(* IEC 61131-3 sources: daoli-st-library/DL_Process (part 36) *)

(* ---- FB_DL_GrateCoolerStartupSeq.st ---- *)
(*
  Name: FB_DL_GrateCoolerStartupSeq
  Category: DL_Process
  Version: 1.0.0
  Round: R91 / 2026-11-25
  开源溯源：clean-room 自研（族 水泥窑篦冷机与预热器，ST 开源生态实测 0 命中，无外部代码引入）
  功能：1) 篦冷机启动序状态机，七相推进：
           待机 → 风机启动 → 篦床低速 → 投料 → 投料升速 → 正常 → （故障）。
           待机相等 xStart 上升沿（必须边沿，防上电即在启动位自动启动）；
           风机相开风机命令并等运行反馈 + 风量达启动下限；篦床低速相给低速指令并等运行反馈；
           投料相开投料命令并等投料反馈；升速相把转速指令按 fRampRpmS 斜率从低速升到正常；
           正常相保持 xDone 并继续风量安全监督，直到 xStart 撤下才回待机。
        2) 每相独立超时 + 整序总超时：相定时器给出正常推进点，相超时定时器给出
           「定时 + DL_OVER_MARGIN」的越限点，整序总超时由 tonTotal 兜底，三者并发监视。
        3) 风量安全监督分两段语义：启动阶段风量不足只拦放行并置信息级码（0121），
           投料之后风量跌破安全下限则进入宽限窗，宽限超时判故障（0128，防篦板过热）。
  边界条件：1) 非有限值闸：风量、转速反馈、周期入参先过 NOT(x > -DL_BIG AND x < DL_BIG)，
           同时拦 NaN 与 Inf；命中即闸断放行（_bAirOk := FALSE / 停机相），
           绝不把 NaN 与 DL_AIR_MIN 比较 —— NaN 比较恒假会伪装成「风量正常」（R19）。
        2) 周期入参闸（R21）：fCycleS <= 0.0 或非有限时，一律改用缺省 DL_CYCLE_DEF = 0.1 s，
           并置信息级码 0129 声明本次斜率按缺省周期折算，不静默。
        3) 时间参数零闸：tFanS / tGrateS / tFeedS / tRampS <= T#0S 时对应相定时器立即置 Q，
           等价于该相跳过（调试用合法组态），语义在此声明，禁上层按「必有停留」假设。
        4) 斜率上限：升速相每拍增量 = fRampRpmS * fCycleS，且指令本身钳在
           [DL_SPD_SLOW, DL_SPD_NORMAL] 内，不用 LIMIT 之后再判超限（R24）。
        5) 故障归因唯一（R190）：风机超时 / 篦床超时 / 投料超时 / 升速超时 / 总超时 /
           外部故障 / 风量不足 / 兜底，八条成因各占独立码值，不共用枚举成员。
        6) 故障解除路径：故障相内 xReset 上升沿 AND NOT xFault AND 入参有限 → 清锁存回待机；
           回待机后必须重新给 xStart 上升沿才能再启动（不自恢复）。
        7) 状态机兜底：CASE 全态覆盖 + ELSE 强制回故障相并置码 0130、清全部输出。
        8) 输出安全初值（R25）：fGrateSpdCmdRpm 初值 0.0（零速为安全侧），
           三个命令位初值 FALSE，待机相显式赋值，防「上电 0 值直穿下发」。
  量纲自证：fRampRpmS 为转速斜率 [rpm/s]，乘 fCycleS [s] 得每拍增量 [rpm]，
           与 fGrateSpdCmdRpm [rpm] 同量纲；fAirFlowNm3h 与 DL_AIR_MIN 同量纲 [Nm3/h]；
           所有时间引脚为 [TIME]，相超时点 = [TIME] + [TIME] = [TIME]，与 TON 的 PT 同量纲。
  码表 Error codes（本件子带 0091_012x，故障级一律 3 行内置 _uFault/_bFault/_eState）:
    16#0091_0121 信息级：风量低于启动下限，风机相暂不放行（不置故障位）
    16#0091_0122 故障级：风机启动超时（定时到但运行反馈未到）
    16#0091_0123 故障级：篦床低速启动超时（无运行反馈）
    16#0091_0124 故障级：投料超时（无投料反馈）
    16#0091_0125 故障级：升速超时（未达正常转速）
    16#0091_0126 故障级：整序总超时
    16#0091_0127 故障级：外部故障输入 xFault
    16#0091_0128 故障级：运行中风量低于安全下限（宽限窗超时）
    16#0091_0129 信息级：周期入参 fCycleS 非法，已按缺省 0.1 s 折算（不置故障位）
    16#0091_0130 故障级：状态机落 ELSE 兜底（非法相位 ID）
    16#0091_0131 故障级：启动序期间风量/转速/斜率入参非有限（NaN 或 Inf）

  修订历史 Revision :
    2026-11-25  v1.0.0  R91 首版
*)

TYPE E_DL_GcsStartupState :
(
    eGcsStartIdle      := 0,    // 待机：等启动上升沿 / Idle, awaiting the start rising edge
    eGcsStartFan       := 10,   // 风机启动：等运行反馈与风量 / Fan start, awaiting feedback and air flow
    eGcsStartSlowGrate := 20,   // 篦床低速：给低速指令等运行反馈 / Grate at low speed, awaiting run feedback
    eGcsStartFeed      := 30,   // 投料：开投料命令等投料反馈 / Feeding, awaiting the feed feedback
    eGcsStartRampUp    := 40,   // 投料升速：按斜率升到正常转速 / Ramping up to normal speed
    eGcsStartNormal    := 50,   // 正常：保持完成位并继续风量监督 / Normal, done held and air supervised
    eGcsStartFault     := 90    // 故障：锁存待解除 / Fault, latched awaiting release
);
END_TYPE

FUNCTION_BLOCK FB_DL_GrateCoolerStartupSeq
VAR_INPUT
    xStart        : BOOL;    // 启动指令（上升沿有效）[bool] / Start command, edge triggered [bool]
    xReset        : BOOL;    // 故障复位（上升沿有效）[bool] / Fault reset, rising edge [bool]
    xFault        : BOOL;    // 外部故障汇总 [bool] / External fault aggregate [bool]
    xFanRunFb     : BOOL;    // 风机运行反馈 [bool] / Fan running feedback [bool]
    xGrateRunFb   : BOOL;    // 篦床驱动运行反馈 [bool] / Grate drive running feedback [bool]
    xFeedRunFb    : BOOL;    // 投料设备运行反馈 [bool] / Feed device running feedback [bool]
    fAirFlowNm3h  : REAL;    // 冷却风量实测值 [Nm3/h] / Measured cooling air flow [Nm3/h]
    fGrateSpdFbRpm : REAL;   // 篦床转速反馈 [rpm] / Grate speed feedback [rpm]
    fRampRpmS     : REAL;    // 升速斜率 [rpm/s] / Speed ramp slope [rpm/s]
    fCycleS       : REAL;    // 任务周期 [s] / Task cycle time [s]
    tFanS         : TIME;    // 风机相设定时长 [TIME] / Fan phase duration [TIME]
    tGrateS       : TIME;    // 篦床低速相设定时长 [TIME] / Low-speed grate phase duration [TIME]
    tFeedS        : TIME;    // 投料相设定时长 [TIME] / Feeding phase duration [TIME]
    tRampS        : TIME;    // 升速相设定时长 [TIME] / Ramp-up phase duration [TIME]
END_VAR
VAR_OUTPUT
    xFanCmd       : BOOL;    // 风机运行命令（安全侧：故障时停）[bool] / Fan run command, fail-safe [bool]
    xGrateCmd     : BOOL;    // 篦床驱动运行命令（安全侧：故障时停）[bool] / Grate drive command, fail-safe [bool]
    xFeedCmd      : BOOL;    // 投料设备运行命令（安全侧：故障时停）[bool] / Feed device command, fail-safe [bool]
    fGrateSpdCmdRpm : REAL;  // 篦床转速指令 [rpm] / Grate speed command [rpm]
    xDone         : BOOL;    // 启动完成保持位 [bool] / Startup complete held flag [bool]
    xBusy         : BOOL;    // 启动进行中 [bool] / Startup sequence busy [bool]
    xAirOk        : BOOL;    // 风量监督通过 [bool] / Air flow supervision passed [bool]
    eState        : E_DL_GcsStartupState;   // 状态出口，段尾单点映射 / State outlet, single-point mapped
    nErrId        : UDINT;   // 事件码，0 = 无事件 / Event code, 0 = none
END_VAR
VAR
    tonFan        : TON;     // 风机相正常定时 [TIME] / Fan phase timer
    tonFanOv      : TON;     // 风机相超时定时 [TIME] / Fan phase overrun timer
    tonGrate      : TON;     // 篦床低速相正常定时 [TIME] / Low-speed grate phase timer
    tonGrateOv    : TON;     // 篦床低速相超时定时 [TIME] / Low-speed grate phase overrun timer
    tonFeed       : TON;     // 投料相正常定时 [TIME] / Feeding phase timer
    tonFeedOv     : TON;     // 投料相超时定时 [TIME] / Feeding phase overrun timer
    tonRamp       : TON;     // 升速相正常定时 [TIME] / Ramp-up phase timer
    tonRampOv     : TON;     // 升速相超时定时 [TIME] / Ramp-up phase overrun timer
    tonTotal      : TON;     // 整序总超时定时 [TIME] / Whole-sequence total timeout timer
    tonAirG       : TON;     // 运行中风量不足宽限定时 [TIME] / Air-shortage grace timer while running
    rtStart       : R_TRIG;  // 启动上升沿检测 [bool] / Start rising edge detector
    rtReset       : R_TRIG;  // 复位上升沿检测 [bool] / Reset rising edge detector
    _eState       : E_DL_GcsStartupState := E_DL_GcsStartupState.eGcsStartIdle;   // 内部相位（CASE 唯一写入目标）
    _eStatePrev   : E_DL_GcsStartupState := E_DL_GcsStartupState.eGcsStartIdle;   // 上一拍相位快照（周期末更新）
    _fSpdSet      : REAL := 0.0;    // 转速指令内部设定值（安全初值零速）[rpm] / Internal speed setpoint, safe init zero [rpm]
    _fCycleUseS   : REAL := 0.1;    // 实际使用的周期值 [s] / Cycle time actually used [s]
    _bFinOk       : BOOL := FALSE;  // 实值入参有限性总闸结果 / Finiteness gate aggregate result
    _bCycleBad    : BOOL := FALSE;  // 周期入参非法标志 [bool] / Cycle input invalid flag [bool]
    _bAirOk       : BOOL := FALSE;  // 风量监督结果 [bool] / Air flow supervision result [bool]
    _bActive      : BOOL := FALSE;  // 启动序激活（风机至正常五相之一）[bool] / Sequence active flag [bool]
    _bRunAirWatch : BOOL := FALSE;  // 投料后风量安全监督生效 [bool] / Post-feed air supervision active [bool]
    _bDoneL       : BOOL := FALSE;  // 完成位锁存（跨相保持）[bool] / Done latch held across phases [bool]
    _bFault       : BOOL := FALSE;  // 故障锁存位 [bool] / Latched fault flag [bool]
    _bRampDone    : BOOL := FALSE;  // 升速到位标志（指令达正常转速）[bool] / Ramp-complete flag [bool]
    _uInfo        : UDINT := 16#0000_0000;   // 信息码，每拍重算 / Info code, recomputed every cycle
    _uFault       : UDINT := 16#0000_0000;   // 故障码锁存 / Latched fault code
    _iPhaseChg    : INT := 0;       // 本拍相位切换计数（观测用）[-] / Phase-change count this cycle [-]
END_VAR
VAR CONSTANT
    DL_EPS        : REAL := 1.0E-9;      // 数值零闸阈值 [-] / Numeric zero gate threshold [-]
    DL_BIG        : REAL := 1.0E12;      // 非有限值闸量级上限 [-] / Finiteness gate magnitude [-]
    DL_CYCLE_DEF  : REAL := 0.1;         // 缺省任务周期 [s] / Default task cycle time [s]
    DL_CYCLE_MIN  : REAL := 0.001;       // 周期合理下限 [s] / Cycle time reasonable low bound [s]
    DL_CYCLE_MAX  : REAL := 10.0;        // 周期合理上限 [s] / Cycle time reasonable high bound [s]
    DL_AIR_MIN    : REAL := 5000.0;      // 启动风量下限 [Nm3/h] / Air flow low limit for start [Nm3/h]
    DL_AIR_SAFE   : REAL := 3000.0;      // 运行风量安全下限 [Nm3/h] / Air flow safety low limit while running [Nm3/h]
    DL_SPD_SLOW   : REAL := 2.0;         // 篦床低速设定 [rpm] / Grate low speed setpoint [rpm]
    DL_SPD_NORMAL : REAL := 12.0;        // 篦床正常转速设定 [rpm] / Grate normal speed setpoint [rpm]
    DL_OVER_MARGIN : TIME := T#30S;      // 相超时相对正常定时的裕量 [TIME] / Phase overrun margin [TIME]
    DL_TOTAL_MAX  : TIME := T#30M;       // 整序总超时上限 [TIME] / Whole-sequence total timeout [TIME]
    DL_AIR_GRACE  : TIME := T#15S;       // 运行中风量不足宽限窗 [TIME] / Air-shortage grace window [TIME]
END_VAR

(* —— 段 0：单拍量预清零（锁存量 _uFault/_bFault/_bDoneL/_eStatePrev 不入清单，R187①） —— *)
_uInfo := 16#0000_0000;                     // 信息码每拍重算 / Info code recomputed
_iPhaseChg := 0;                            // 相位切换计数每拍重算 / Phase-change counter recomputed
nErrId := 16#0000_0000;                     // 事件码缺省无事件 / Event code defaults to none

(* —— 段 1：周期入参闸（R21：非法周期不静默，改用缺省并置信息码） —— *)
_bCycleBad := NOT (fCycleS > -DL_BIG AND fCycleS < DL_BIG)
              OR (fCycleS < DL_CYCLE_MIN) OR (fCycleS > DL_CYCLE_MAX);
IF _bCycleBad THEN
    _fCycleUseS := DL_CYCLE_DEF;            // 非法周期一律用缺省 0.1 s
    _uInfo := 16#0091_0129;                 // 信息级：周期入参非法，已用缺省（不置故障位）
ELSE
    _fCycleUseS := fCycleS;                 // 合法周期原值使用
END_IF

(* —— 段 2：非有限值闸（R19：闸断实值通路，风量/转速/斜率任一非有限即拒绝放行） —— *)
_bFinOk := (fAirFlowNm3h > -DL_BIG) AND (fAirFlowNm3h < DL_BIG)
           AND (fGrateSpdFbRpm > -DL_BIG) AND (fGrateSpdFbRpm < DL_BIG)
           AND (fRampRpmS > -DL_BIG) AND (fRampRpmS < DL_BIG);

(* —— 段 3：风量监督（启动用下限；非有限值直接判不通过，不参与比较） —— *)
IF NOT _bFinOk THEN
    _bAirOk := FALSE;                       // 非有限一律判不通过（安全侧）
ELSE
    _bAirOk := (fAirFlowNm3h >= DL_AIR_MIN);
END_IF

(* —— 段 4：状态派生量（本拍相位为上一拍末值，标准 FB 周期语义） —— *)
_bActive := (_eState = E_DL_GcsStartupState.eGcsStartFan)
            OR (_eState = E_DL_GcsStartupState.eGcsStartSlowGrate)
            OR (_eState = E_DL_GcsStartupState.eGcsStartFeed)
            OR (_eState = E_DL_GcsStartupState.eGcsStartRampUp)
            OR (_eState = E_DL_GcsStartupState.eGcsStartNormal);
_bRunAirWatch := (_eState = E_DL_GcsStartupState.eGcsStartFeed)
                 OR (_eState = E_DL_GcsStartupState.eGcsStartRampUp)
                 OR (_eState = E_DL_GcsStartupState.eGcsStartNormal);

(* —— 段 5：定时器与边沿无条件周期刷新（R7：调用语句不得置于 IF/CASE 内） —— *)
rtStart(CLK := xStart);                                                                 // 启动上升沿，每拍必调
rtReset(CLK := xReset);                                                                 // 复位上升沿，每拍必调
tonFan(IN := (_eState = E_DL_GcsStartupState.eGcsStartFan), PT := tFanS);               // 风机相正常定时
tonFanOv(IN := (_eState = E_DL_GcsStartupState.eGcsStartFan), PT := tFanS + DL_OVER_MARGIN);      // 风机相超时点
tonGrate(IN := (_eState = E_DL_GcsStartupState.eGcsStartSlowGrate), PT := tGrateS);     // 篦床低速相正常定时
tonGrateOv(IN := (_eState = E_DL_GcsStartupState.eGcsStartSlowGrate),
           PT := tGrateS + DL_OVER_MARGIN);                                             // 篦床低速相超时点
tonFeed(IN := (_eState = E_DL_GcsStartupState.eGcsStartFeed), PT := tFeedS);            // 投料相正常定时
tonFeedOv(IN := (_eState = E_DL_GcsStartupState.eGcsStartFeed), PT := tFeedS + DL_OVER_MARGIN);   // 投料相超时点
tonRamp(IN := (_eState = E_DL_GcsStartupState.eGcsStartRampUp), PT := tRampS);          // 升速相正常定时
tonRampOv(IN := (_eState = E_DL_GcsStartupState.eGcsStartRampUp), PT := tRampS + DL_OVER_MARGIN); // 升速相超时点
tonTotal(IN := _bActive, PT := DL_TOTAL_MAX);                                           // 整序总超时
tonAirG(IN := _bRunAirWatch AND (NOT _bAirOk) AND (NOT _bFault), PT := DL_AIR_GRACE);    // 风量不足宽限窗

(* —— 段 6：全局故障拦截（优先级最高；已锁存则不再改写码值，禁同拍抹除） —— *)
IF xFault AND (NOT _bFault) THEN
    _uFault := 16#0091_0127;                // 故障级：外部故障输入
    _bFault := TRUE;                        // 锁存（3 行内置，R45 配对）
    _eState := E_DL_GcsStartupState.eGcsStartFault;
END_IF
IF tonTotal.Q AND _bActive AND (NOT _bFault) THEN
    _uFault := 16#0091_0126;                // 故障级：整序总超时
    _bFault := TRUE;                        // 锁存
    _eState := E_DL_GcsStartupState.eGcsStartFault;
END_IF
IF tonAirG.Q AND (NOT _bFault) THEN
    _uFault := 16#0091_0128;                // 故障级：运行中风量低于安全下限
    _bFault := TRUE;                        // 锁存
    _eState := E_DL_GcsStartupState.eGcsStartFault;
END_IF
IF (NOT _bFinOk) AND (NOT _bFault) AND _bActive THEN
    _uFault := 16#0091_0131;                // 故障级：启动序期间入参非有限（独立成因，不与风机超时共用码）
    _bFault := TRUE;                        // 锁存
    _eState := E_DL_GcsStartupState.eGcsStartFault;
END_IF

(* —— 段 7：相位机（只做迁移与内部状态更新；出口在段 9 单点映射） —— *)
CASE _eState OF

E_DL_GcsStartupState.eGcsStartIdle:
    _fSpdSet := 0.0;                        // 待机转速指令显式零（安全侧，R25）
    _bRampDone := FALSE;                    // 待机重置升速到位标志
    IF NOT xStart THEN
        _bDoneL := FALSE;                   // 撤令即清完成位，为下次启动重新武装
    ELSIF NOT _bAirOk THEN
        _uInfo := 16#0091_0121;             // 信息级：风量不足，风机相暂不放行
    ELSIF rtStart.Q THEN
        _bDoneL := FALSE;                   // 新序开始：清完成位（迁移前一次性清）
        _eState := E_DL_GcsStartupState.eGcsStartFan;   // 进风机启动相
    END_IF

E_DL_GcsStartupState.eGcsStartFan:
    IF NOT xStart THEN
        _uFault := 16#0091_0127;            // 故障级：启动中撤令，按外部中断归因
        _bFault := TRUE;                    // 锁存
        _eState := E_DL_GcsStartupState.eGcsStartFault;
    ELSIF tonFanOv.Q THEN
        _uFault := 16#0091_0122;            // 故障级：风机启动超时
        _bFault := TRUE;                    // 锁存
        _eState := E_DL_GcsStartupState.eGcsStartFault;
    ELSIF tonFan.Q AND xFanRunFb AND _bAirOk THEN
        _eState := E_DL_GcsStartupState.eGcsStartSlowGrate;   // 本拍合法事件优先于超时迁移（R275）
    ELSE
        _uInfo := 16#0091_0121;             // 信息级：风量/反馈未就绪，继续等
    END_IF

E_DL_GcsStartupState.eGcsStartSlowGrate:
    _fSpdSet := DL_SPD_SLOW;                // 低速相：转速指令置低速设定
    IF NOT xStart THEN
        _uFault := 16#0091_0127;            // 故障级：启动中撤令
        _bFault := TRUE;                    // 锁存
        _eState := E_DL_GcsStartupState.eGcsStartFault;
    ELSIF tonGrateOv.Q THEN
        _uFault := 16#0091_0123;            // 故障级：篦床低速启动超时
        _bFault := TRUE;                    // 锁存
        _eState := E_DL_GcsStartupState.eGcsStartFault;
    ELSIF tonGrate.Q AND xGrateRunFb THEN
        _eState := E_DL_GcsStartupState.eGcsStartFeed;        // 进投料相
    END_IF

E_DL_GcsStartupState.eGcsStartFeed:
    _fSpdSet := DL_SPD_SLOW;                // 投料相：转速保持低速
    IF NOT xStart THEN
        _uFault := 16#0091_0127;            // 故障级：投料中撤令
        _bFault := TRUE;                    // 锁存
        _eState := E_DL_GcsStartupState.eGcsStartFault;
    ELSIF tonFeedOv.Q THEN
        _uFault := 16#0091_0124;            // 故障级：投料超时
        _bFault := TRUE;                    // 锁存
        _eState := E_DL_GcsStartupState.eGcsStartFault;
    ELSIF tonFeed.Q AND xFeedRunFb THEN
        _eState := E_DL_GcsStartupState.eGcsStartRampUp;      // 进升速相
    END_IF

E_DL_GcsStartupState.eGcsStartRampUp:
    _fSpdSet := LIMIT(DL_SPD_SLOW, _fSpdSet + fRampRpmS * _fCycleUseS, DL_SPD_NORMAL);   // 每拍按斜率升速
    _bRampDone := (_fSpdSet >= DL_SPD_NORMAL);                                            // 到位判据（用钳后设定值即可）
    IF NOT xStart THEN
        _uFault := 16#0091_0127;            // 故障级：升速中撤令
        _bFault := TRUE;                    // 锁存
        _eState := E_DL_GcsStartupState.eGcsStartFault;
    ELSIF tonRampOv.Q AND (NOT _bRampDone) THEN
        _uFault := 16#0091_0125;            // 故障级：升速超时
        _bFault := TRUE;                    // 锁存
        _eState := E_DL_GcsStartupState.eGcsStartFault;
    ELSIF _bRampDone AND tonRamp.Q THEN
        _bDoneL := TRUE;                    // 完成位锁存（跨相保持，段 9 单点映射）
        _eState := E_DL_GcsStartupState.eGcsStartNormal;      // 进正常相
    END_IF

E_DL_GcsStartupState.eGcsStartNormal:
    _fSpdSet := DL_SPD_NORMAL;              // 正常相：转速指令置正常设定
    IF NOT xStart THEN
        _bDoneL := FALSE;                   // 撤令：清完成位并回待机（命令随之撤销）
        _bRampDone := FALSE;                // 升速标志一并清，下次重新走斜率
        _eState := E_DL_GcsStartupState.eGcsStartIdle;
    ELSIF NOT _bAirOk THEN
        _uInfo := 16#0091_0121;             // 信息级：风量偏低但仍在宽限窗内（宽限超时由段 6 判故障）
    END_IF

E_DL_GcsStartupState.eGcsStartFault:
    _fSpdSet := 0.0;                        // 故障相转速指令强制零（安全侧，R25）
    IF rtReset.Q AND (NOT xFault) AND _bFinOk THEN
        _bFault := FALSE;                   // 解除路径：复位沿 + 外部故障消失 + 入参有限（可达，R188）
        _uFault := 16#0000_0000;            // 清锁存码
        _bDoneL := FALSE;                   // 完成位一并清，避免故障后误报完成
        _bRampDone := FALSE;                // 升速标志清，需重新走完整序
        _eState := E_DL_GcsStartupState.eGcsStartIdle;        // 回待机，需新上升沿才可再启动
    END_IF

ELSE
    _uFault := 16#0091_0130;                // 故障级：非法相位 ID 兜底
    _bFault := TRUE;                        // 锁存
    _fSpdSet := 0.0;                        // 兜底侧转速强制零
    _eState := E_DL_GcsStartupState.eGcsStartFault;           // 强制回故障相

END_CASE

(* —— 段 8：后置段（相位快照在迁移判断之后统一更新） —— *)
IF _eState <> _eStatePrev THEN
    _iPhaseChg := _iPhaseChg + 1;           // 相位已切换：记一拍切换事件（观测用）
END_IF
_eStatePrev := _eState;                     // 快照在周期末尾统一更新

(* —— 段 9：出口单点映射（名实同源；命令由状态导出，故障侧一律撤销） —— *)
xFanCmd := ((_eState = E_DL_GcsStartupState.eGcsStartFan)
            OR (_eState = E_DL_GcsStartupState.eGcsStartSlowGrate)
            OR (_eState = E_DL_GcsStartupState.eGcsStartFeed)
            OR (_eState = E_DL_GcsStartupState.eGcsStartRampUp)
            OR (_eState = E_DL_GcsStartupState.eGcsStartNormal)) AND (NOT _bFault);        // 风机：五相开
xGrateCmd := ((_eState = E_DL_GcsStartupState.eGcsStartSlowGrate)
              OR (_eState = E_DL_GcsStartupState.eGcsStartFeed)
              OR (_eState = E_DL_GcsStartupState.eGcsStartRampUp)
              OR (_eState = E_DL_GcsStartupState.eGcsStartNormal)) AND (NOT _bFault);      // 篦床：四相开
xFeedCmd := ((_eState = E_DL_GcsStartupState.eGcsStartFeed)
             OR (_eState = E_DL_GcsStartupState.eGcsStartRampUp)
             OR (_eState = E_DL_GcsStartupState.eGcsStartNormal)) AND (NOT _bFault);       // 投料：三相开
IF xGrateCmd THEN
    fGrateSpdCmdRpm := _fSpdSet;            // 转速指令出口（单点写，分支互斥）
ELSE
    fGrateSpdCmdRpm := 0.0;                 // 未开篦床即零速指令（安全侧，R25）
END_IF
xDone := _bDoneL AND (NOT _bFault);                                        // 完成位出口
xBusy := _bActive AND (NOT _bFault);                                       // 进行中出口
xAirOk := _bAirOk;                                                         // 风量监督出口
eState := _eState;                                                         // 状态出口单点映射
IF _bFault THEN
    nErrId := _uFault;                      // 故障锁存码回放（不在故障相按当下输入重推断）
ELSE
    nErrId := _uInfo;                       // 信息码
END_IF

END_FUNCTION_BLOCK

(* ---- FB_DL_GrateCoolerStrokeWatch.st ---- *)
(*
  Name: FB_DL_GrateCoolerStrokeWatch
  Category: DL_Process
  Version: 1.0.0
  Round: R91 / 2026-11-25
  开源溯源：clean-room 自研（族 水泥窑篦冷机与预热器，ST 开源生态实测 0 命中，无外部代码引入）
  功能：1) 篦床行程三判据并行监视，各自独立去抖：
           ① 行程超限：MAX(左/右行程) > fStrokeMaxMm（篦板越程会顶死液压缸）；
           ② 左右不同步：|左 − 右| > fSyncMaxMm（双侧不同步导致篦床歪斜与卡阻）；
           ③ 停滞：有运行指令 xEnable 且一个去抖窗内位移 < DL_MOVE_EPS（液压失压或机械卡死）。
        2) 三级报警升级：原始判据成立即进预警相（信息级码）；去抖确认后单成因进报警相（故障级码，
           不直接停机）；两成因及以上并发进停机建议相（最高级码，建议上层连锁停机）。
        3) 锁存与解除：报警相与停机建议相的故障码一律锁存回放，唯一解除路径为 xReset 上升沿，
           且解除时必须「三判据原始值全部消失」才回正常相（防止带病复位后立刻再报）。
  边界条件：1) 非有限值闸：五路实值入参先过 NOT(x > -DL_BIG AND x < DL_BIG)，同时拦 NaN 与 Inf；
           命中即置故障锁存（码 0117）并进故障相，而不是把 NaN 拿去与限值比较 ——
           NaN 比较恒假会把「测点断线」伪装成「行程正常」（R19）。
        2) 组态域闸：fStrokeMaxMm / fSyncMaxMm 必须 > DL_EPS，tDebounce / tStallS 必须 > T#0S，
           越域置码 0118 并进故障相（去抖窗为零会让判据无滞后直达停机）。
        3) 位移快照闸：首拍 _bPrevValid = FALSE 时不判停滞，避免上电首个扫描周期
           「上拍行程 = 0」造成的假停滞。
        4) 定时器周期刷新（R7）：四个 TON 实例全部在 CASE 之外无条件调用，IN 由状态与判据导出，
           相迁移即 IN 归假自复位，不靠外部沿清零（R188）。
        5) 状态机兜底：CASE 全态覆盖 + ELSE 强制进故障相并置码 0116、清全部输出。
        6) 输出安全初值（R25）：xWarn / xAlarm / xStopSuggest 初值 FALSE，nLevel 初值 0，
           待机相显式赋值，防「上电未初始化直穿」。
  量纲自证：fStrokeLeftMm / fStrokeRightMm / fStrokeMaxMm / fSyncMaxMm 均为长度 [mm]，
           比较两侧同量纲；位移差 |左 − 右| 仍为 [mm]；
           tDebounce / tStallS 为 [TIME]，直接作为 TON 的 PT，无跨量纲运算。
  码表 Error codes（本件子带 0091_011x，故障级一律 3 行内置 _uFault/_bFault/_eState）:
    16#0091_0111 信息级：行程判据预警（原始值成立，尚在去抖窗内，不置故障位）
    16#0091_0112 故障级：左侧行程超限（去抖确认）
    16#0091_0113 故障级：左右行程不同步（去抖确认）
    16#0091_0114 故障级：篦床停滞，有运行指令但无位移（去抖确认）
    16#0091_0115 故障级：两成因及以上并发，建议停机
    16#0091_0116 故障级：状态机落 ELSE 兜底（非法相位 ID）
    16#0091_0117 故障级：行程或限值入参非有限（NaN / Inf）
    16#0091_0118 故障级：组态越域（行程限值或去抖窗为零/为负）

  修订历史 Revision :
    2026-11-25  v1.0.0  R91 首版
*)

TYPE E_DL_GcsStrokeWatchState :
(
    eGcsStrokeNormal := 0,    // 正常：三判据原始值全部消失 / Normal, all three raw criteria cleared
    eGcsStrokeWarn   := 10,   // 预警：原始判据成立，等去抖窗 / Warning, raw criterion present, debounce running
    eGcsStrokeAlarm  := 20,   // 报警：单成因去抖确认，锁存待复位 / Alarm, single cause confirmed and latched
    eGcsStrokeTrip   := 30,   // 停机建议：两成因及以上并发 / Trip advice, two or more causes together
    eGcsStrokeFault  := 90    // 故障：入参/组态非法，锁存待复位 / Fault, invalid input or configuration, latched
);
END_TYPE

FUNCTION_BLOCK FB_DL_GrateCoolerStrokeWatch
VAR_INPUT
    xEnable        : BOOL;    // 监视使能（篦床运行指令）[bool] / Monitoring enable, grate run command [bool]
    xReset         : BOOL;    // 故障复位（上升沿有效）[bool] / Fault reset, rising edge [bool]
    xFault         : BOOL;    // 外部故障汇总 [bool] / External fault aggregate [bool]
    fStrokeLeftMm  : REAL;    // 左侧油缸行程 [mm] / Left cylinder stroke [mm]
    fStrokeRightMm : REAL;    // 右侧油缸行程 [mm] / Right cylinder stroke [mm]
    fStrokeMaxMm   : REAL;    // 允许最大行程 [mm] / Permitted maximum stroke [mm]
    fSyncMaxMm     : REAL;    // 左右允许最大行程差 [mm] / Permitted maximum stroke difference [mm]
    tDebounce      : TIME;    // 判据去抖窗 [TIME] / Criteria debounce window [TIME]
    tStallS        : TIME;    // 停滞判定窗 [TIME] / Stall detection window [TIME]
END_VAR
VAR_OUTPUT
    xWarn          : BOOL;    // 预警位（信息级）[bool] / Warning flag, information grade [bool]
    xAlarm         : BOOL;    // 报警位（故障级）[bool] / Alarm flag, fault grade [bool]
    xStopSuggest   : BOOL;    // 停机建议位 [bool] / Stop suggestion flag [bool]
    nLevel         : INT;     // 报警等级 0=正常 1=预警 2=报警 3=停机 [level] / Alarm level 0..3 [level]
    eState         : E_DL_GcsStrokeWatchState;   // 状态出口，段尾单点映射 / State outlet, single-point mapped
    nErrId         : UDINT;   // 事件码，0 = 无事件 / Event code, 0 = none
END_VAR
VAR
    tonOver        : TON;     // 行程超限去抖定时 [TIME] / Stroke-overrun debounce timer
    tonSync        : TON;     // 左右不同步去抖定时 [TIME] / Synchronism debounce timer
    tonStall       : TON;     // 停滞判定定时 [TIME] / Stall detection timer
    tonClear       : TON;     // 复位清障确认定时 [TIME] / Reset clearance confirmation timer
    rtReset        : R_TRIG;  // 复位上升沿检测 [bool] / Reset rising edge detector
    _eState        : E_DL_GcsStrokeWatchState := E_DL_GcsStrokeWatchState.eGcsStrokeNormal;   // 内部相位（CASE 唯一写入目标）
    _fStrokePrevMm : REAL := 0.0;   // 上拍左侧行程快照 [mm] / Previous-cycle left stroke snapshot [mm]
    _bPrevValid    : BOOL := FALSE; // 行程快照有效位（首拍为假）/ Stroke snapshot validity, false on first cycle
    _bFinOk        : BOOL := FALSE; // 实值入参有限性总闸结果 / Finiteness gate aggregate result
    _bCfgOk        : BOOL := FALSE; // 组态参数域闸结果 / Configuration domain gate result
    _bOverRaw      : BOOL := FALSE; // 行程超限原始判据 [bool] / Raw stroke-overrun criterion
    _bSyncRaw      : BOOL := FALSE; // 左右不同步原始判据 [bool] / Raw synchronism criterion
    _bStallRaw     : BOOL := FALSE; // 停滞原始判据 [bool] / Raw stall criterion
    _bAnyRaw       : BOOL := FALSE; // 三判据任一成立 [bool] / Any raw criterion present
    _iCauseNum     : INT := 0;      // 已去抖确认的成因数 [-]/ Confirmed cause count [-]
    _bAlarmL       : BOOL := FALSE; // 报警锁存位 [bool] / Latched alarm flag
    _bTripL        : BOOL := FALSE; // 停机建议锁存位 [bool] / Latched trip-advice flag
    _bFault        : BOOL := FALSE; // 故障锁存位 [bool] / Latched fault flag
    _uInfo         : UDINT := 16#0000_0000;   // 信息码，每拍重算 / Info code, recomputed every cycle
    _uFault        : UDINT := 16#0000_0000;   // 故障码锁存 / Latched fault code
END_VAR
VAR CONSTANT
    DL_EPS         : REAL := 1.0E-9;    // 数值零闸阈值 [-] / Numeric zero gate threshold [-]
    DL_BIG         : REAL := 1.0E12;    // 非有限值闸量级上限 [-] / Finiteness gate magnitude [-]
    DL_MOVE_EPS    : REAL := 0.05;      // 判定「有位移」的最小行程变化 [mm] / Minimum movement to count as moving [mm]
    DL_ZERO_MM     : REAL := 0.0;       // 行程零基准 [mm] / Zero stroke reference [mm]
    DL_CLEAR_CHK   : TIME := T#3S;      // 复位清障确认窗 [TIME] / Reset clearance confirmation window [TIME]
END_VAR

(* —— 段 0：单拍量预清零（锁存量 _uFault/_bFault/_bAlarmL/_bTripL 不入清单，R187①） —— *)
_uInfo := 16#0000_0000;                     // 信息码每拍重算 / Info code recomputed
nErrId := 16#0000_0000;                     // 事件码缺省无事件 / Event code defaults to none
_iCauseNum := 0;                            // 成因计数每拍重算 / Cause counter recomputed

(* —— 段 1：非有限值闸与组态域闸（R19：不拿 NaN 去比较，直接判故障） —— *)
_bFinOk := (fStrokeLeftMm > -DL_BIG) AND (fStrokeLeftMm < DL_BIG)
           AND (fStrokeRightMm > -DL_BIG) AND (fStrokeRightMm < DL_BIG)
           AND (fStrokeMaxMm > -DL_BIG) AND (fStrokeMaxMm < DL_BIG)
           AND (fSyncMaxMm > -DL_BIG) AND (fSyncMaxMm < DL_BIG);
_bCfgOk := (fStrokeMaxMm > DL_EPS)          // 行程限值必须为正
           AND (fSyncMaxMm > DL_EPS)        // 同步差限值必须为正
           AND (tDebounce > T#0S)           // 去抖窗必须为正
           AND (tStallS > T#0S);            // 停滞窗必须为正

(* —— 段 2：判据派生（原始值；LIMIT 不参与，避免判据恒真，R24） —— *)
_bOverRaw := _bFinOk AND _bCfgOk
             AND ((MAX(fStrokeLeftMm, fStrokeRightMm) > fStrokeMaxMm)
                  OR (MIN(fStrokeLeftMm, fStrokeRightMm) < DL_ZERO_MM));
_bSyncRaw := _bFinOk AND _bCfgOk
             AND (ABS(fStrokeLeftMm - fStrokeRightMm) > fSyncMaxMm);
_bStallRaw := _bFinOk AND _bCfgOk AND xEnable AND _bPrevValid
              AND (ABS(fStrokeLeftMm - _fStrokePrevMm) < DL_MOVE_EPS);
_bAnyRaw := _bOverRaw OR _bSyncRaw OR _bStallRaw;

(* —— 段 3：定时器与边沿无条件周期刷新（R7：调用语句不得置于 IF/CASE 内） —— *)
rtReset(CLK := xReset);                                                     // 复位上升沿，每拍必调
tonOver(IN := _bOverRaw AND (NOT _bFault), PT := tDebounce);                 // 行程超限去抖
tonSync(IN := _bSyncRaw AND (NOT _bFault), PT := tDebounce);                 // 同步差去抖
tonStall(IN := _bStallRaw AND (NOT _bFault), PT := tStallS);                 // 停滞判定
tonClear(IN := rtReset.Q, PT := DL_CLEAR_CHK);                               // 复位清障确认，自复位靠 rtReset 单拍

(* —— 段 4：相位机（只做迁移与锁存；出口在段 6 单点映射） —— *)
CASE _eState OF

E_DL_GcsStrokeWatchState.eGcsStrokeNormal:
    IF (NOT _bFinOk) OR (NOT _bCfgOk) THEN
        IF NOT _bFinOk THEN
            _uFault := 16#0091_0117;        // 故障级：入参非有限（唯一归因，R190）
        ELSE
            _uFault := 16#0091_0118;        // 故障级：组态越域（唯一归因，R190）
        END_IF
        _bFault := TRUE;                    // 锁存（3 行内置，R45 配对）
        _bAlarmL := FALSE;                  // 报警锁存清，避免双码并存
        _bTripL := FALSE;                   // 停机建议锁存清
        _eState := E_DL_GcsStrokeWatchState.eGcsStrokeFault;
    ELSIF xFault THEN
        _uFault := 16#0091_0115;            // 故障级：外部故障按最高级归因（由上层提供）
        _bFault := TRUE;                    // 锁存
        _bAlarmL := FALSE;                  // 报警锁存清
        _bTripL := FALSE;                   // 停机建议锁存清
        _eState := E_DL_GcsStrokeWatchState.eGcsStrokeFault;
    ELSIF _bAnyRaw THEN
        _eState := E_DL_GcsStrokeWatchState.eGcsStrokeWarn;   // 原始判据成立：进预警相等去抖
    END_IF

E_DL_GcsStrokeWatchState.eGcsStrokeWarn:
    IF tonOver.Q THEN
        _iCauseNum := _iCauseNum + 1;       // 成因 1：行程超限已确认
    END_IF
    IF tonSync.Q THEN
        _iCauseNum := _iCauseNum + 1;       // 成因 2：不同步已确认
    END_IF
    IF tonStall.Q THEN
        _iCauseNum := _iCauseNum + 1;       // 成因 3：停滞已确认
    END_IF
    IF _iCauseNum >= 2 THEN
        _uFault := 16#0091_0115;            // 故障级：两成因及以上并发，建议停机
        _bTripL := TRUE;                    // 停机建议锁存
        _eState := E_DL_GcsStrokeWatchState.eGcsStrokeTrip;
    ELSIF tonOver.Q THEN
        _uFault := 16#0091_0112;            // 故障级：左侧/最高侧行程超限
        _bAlarmL := TRUE;                   // 报警锁存
        _eState := E_DL_GcsStrokeWatchState.eGcsStrokeAlarm;
    ELSIF tonSync.Q THEN
        _uFault := 16#0091_0113;            // 故障级：左右行程不同步
        _bAlarmL := TRUE;                   // 报警锁存
        _eState := E_DL_GcsStrokeWatchState.eGcsStrokeAlarm;
    ELSIF tonStall.Q THEN
        _uFault := 16#0091_0114;            // 故障级：篦床停滞
        _bAlarmL := TRUE;                   // 报警锁存
        _eState := E_DL_GcsStrokeWatchState.eGcsStrokeAlarm;
    ELSIF NOT _bAnyRaw THEN
        _eState := E_DL_GcsStrokeWatchState.eGcsStrokeNormal;   // 判据自行消失：回正常，不留痕
    ELSE
        _uInfo := 16#0091_0111;             // 信息级：预警中（尚在去抖窗内，不置故障位）
    END_IF

E_DL_GcsStrokeWatchState.eGcsStrokeAlarm:
    IF rtReset.Q THEN
        _bAlarmL := FALSE;                  // 解除路径：复位上升沿（可达，R188）
        _uFault := 16#0000_0000;            // 清锁存码
        _eState := E_DL_GcsStrokeWatchState.eGcsStrokeNormal;
    END_IF

E_DL_GcsStrokeWatchState.eGcsStrokeTrip:
    IF rtReset.Q THEN
        _bTripL := FALSE;                   // 解除路径：复位上升沿（可达，R188）
        _uFault := 16#0000_0000;            // 清锁存码
        _eState := E_DL_GcsStrokeWatchState.eGcsStrokeNormal;
    END_IF

E_DL_GcsStrokeWatchState.eGcsStrokeFault:
    IF rtReset.Q AND (NOT xFault) AND _bFinOk AND _bCfgOk THEN
        _bFault := FALSE;                   // 解除路径：复位沿 + 外部故障消失 + 入参与组态合法（可达）
        _uFault := 16#0000_0000;            // 清锁存码
        _eState := E_DL_GcsStrokeWatchState.eGcsStrokeNormal;
    END_IF

ELSE
    _uFault := 16#0091_0116;                // 故障级：非法相位 ID 兜底
    _bFault := TRUE;                        // 锁存
    _bAlarmL := FALSE;                      // 报警锁存清
    _bTripL := FALSE;                       // 停机建议锁存清
    _eState := E_DL_GcsStrokeWatchState.eGcsStrokeFault;   // 强制回故障相

END_CASE

(* —— 段 5：后置段（行程快照在迁移判断之后统一更新，禁在分支内散写） —— *)
IF _bFinOk THEN
    _fStrokePrevMm := fStrokeLeftMm;        // 快照更新（仅有限值可信时才更新）
    _bPrevValid := TRUE;                    // 快照自此有效
ELSE
    _bPrevValid := FALSE;                   // 非有限值使快照失效，防污染下一拍停滞判据
END_IF

(* —— 段 6：出口单点映射（名实同源；故障与锁存位一律由状态导出） —— *)
xWarn := (_eState = E_DL_GcsStrokeWatchState.eGcsStrokeWarn);                          // 预警仅预警相
xAlarm := _bAlarmL AND (NOT _bFault) AND (NOT _bTripL);                                // 报警：锁存且未升级
xStopSuggest := _bTripL OR _bFault;                                                    // 停机建议：并发或故障相
IF _bTripL OR _bFault THEN
    nLevel := 3;                            // 最高级：停机建议
ELSIF _bAlarmL THEN
    nLevel := 2;                            // 报警级
ELSIF xWarn THEN
    nLevel := 1;                            // 预警级
ELSE
    nLevel := 0;                            // 正常
END_IF
eState := _eState;                          // 状态出口单点映射
IF _bTripL OR _bFault OR _bAlarmL THEN
    nErrId := _uFault;                      // 故障码锁存回放（不在故障相按当下输入重推断）
ELSE
    nErrId := _uInfo;                       // 信息码（预警中）
END_IF

END_FUNCTION_BLOCK

(* ---- FB_DL_HandAutoModeGateBank.st ---- *)
//==============================================================================
// 功能块：FB_DL_HandAutoModeGateBank ｜ 中文名称：手/自动模式权限门组（双钥匙）
// 所属子库：DL_Process ｜ 版本：v1.0.0 ｜ 日期：2026-11-23
// 兼容：CODESYS V3.5+ / TwinCAT 3 / 汇川 InoProShop（纯 IEC 61131-3，零方言）
// 功能描述：2 回路手/自动模式权限门 Bank：模式切换须"双钥匙同时确认"
//           （bKeyA AND bKeyB）+ 模式请求沿，双钥匙缺一拒绝切换（信息级
//           留痕）。模式切换沿经审计计数器（UDINT 饱和不回绕）留痕，供
//           ISA-88/PackML 相语义审计。两回路逻辑同构独立驻留。
// 开源溯源 (Origin)：候选队列 MANUAL（oscatBasic，MIT 许可，
//           https://github.com/tkucic/brOscatLib/blob/main/oscatBasic/MANUAL.st）
//           与 CONTROL_MODE（AixOCAT，MIT 许可，
//           https://github.com/RWTH-EBC/AixOCAT/blob/develop/OSCAT/OSCAT/OSCAT/oscat_basic/Data%20types/CONTROL_MODE.TcDUT）
//           ——手/自动模式选择与模式枚举行为定义参考；原名 MANUAL /
//           CONTROL_MODE → 道莅 FB_DL_HandAutoModeGateBank，clean-room
//           独立重写（双钥匙确认 + 沿审计为道莅增量，零源码行复制）
// 公开接口清单：输入 {bAutoReq1/2, bManReq1/2, bKeyA1/2, bKeyB1/2}；
//               输出 {eMode1/2, bSwitchPulse1/2, uAuditCnt1/2} / uErrCode / bValid
// 错误码表：16#0005_3060 信息级（回路 1 单钥匙拒绝切换，不置 bError）/
//           16#0005_3061 信息级（回路 2 单钥匙拒绝切换，不置 bError）/
//           16#0005_3062 信息级（审计计数饱和不回绕，不置 bError）/
//           16#0005_3063 预留禁用（不得挪用）
// 状态机：E_DL_HaMode（本文件唯一定义，全库唯一属主）：
//           eAuto = 0 / eManual = 1；非法模式值走 CASE ELSE 兜底归 eManual
//           （人工介入侧为安全侧）
// 边界行为：① 双钥匙缺一切换请求沿 → 拒绝 + 信息码（不切换）；
//           ② 切换成功拍发单拍脉冲 bSwitchPulse（两段式出口映射）；
//           ③ 审计计数饱和于 4294967295 不回绕（信息级留痕）；
//           ④ R_TRIG ×8 每拍无条件刷新（不入分支，红线 R7）；
//           ⑤ CASE 带 ELSE 非法模式兜底归 eManual。
// 修订历史：v1.0.0 2026-11-23 首版（R73 派单 · 批 2 · 序 19）
//==============================================================================

(*------------------------------------------------------------------------------
 * 枚举: E_DL_HaMode（归属本功能块，同文件发布，全库唯一属主）
 * 含义: 手/自动模式，成员与 CASE 标签双向完备。
 *-----------------------------------------------------------------------------*)
TYPE E_DL_HaMode :
(
    eAuto   := 0,   // 自动模式：上层顺控驱动 / Auto mode, driven by the upper sequence
    eManual := 1    // 手动模式：操作员直接驱动 / Manual mode, operator direct drive
);
END_TYPE

(*==============================================================================
 * 功能块: FB_DL_HandAutoModeGateBank
 * 调用约定: 每个扫描周期无条件调用一次；实例状态全部驻留于私有变量。
 *==============================================================================*)
FUNCTION_BLOCK FB_DL_HandAutoModeGateBank
VAR_INPUT
    bAutoReq1 : BOOL := FALSE;         // 回路 1 自动请求（沿触发）/ Loop 1 auto request, edge triggered
    bManReq1  : BOOL := FALSE;         // 回路 1 手动请求（沿触发）/ Loop 1 manual request, edge triggered
    bKeyA1    : BOOL := FALSE;         // 回路 1 钥匙 A（切换期须保持）/ Loop 1 key A, held during switching
    bKeyB1    : BOOL := FALSE;         // 回路 1 钥匙 B（切换期须保持）/ Loop 1 key B, held during switching
    bAutoReq2 : BOOL := FALSE;         // 回路 2 自动请求（沿触发）/ Loop 2 auto request, edge triggered
    bManReq2  : BOOL := FALSE;         // 回路 2 手动请求（沿触发）/ Loop 2 manual request, edge triggered
    bKeyA2    : BOOL := FALSE;         // 回路 2 钥匙 A（切换期须保持）/ Loop 2 key A, held during switching
    bKeyB2    : BOOL := FALSE;         // 回路 2 钥匙 B（切换期须保持）/ Loop 2 key B, held during switching
END_VAR
VAR_OUTPUT
    eMode1    : E_DL_HaMode;           // 回路 1 当前模式 / Loop 1 current mode
    eMode2    : E_DL_HaMode;           // 回路 2 当前模式 / Loop 2 current mode
    bSwitchPulse1 : BOOL;              // 回路 1 单拍切换脉冲 / Loop 1 single-scan switch pulse
    bSwitchPulse2 : BOOL;              // 回路 2 单拍切换脉冲 / Loop 2 single-scan switch pulse
    uAuditCnt1: UDINT;                 // 回路 1 模式切换审计计数 [次] / Loop 1 switch audit count
    uAuditCnt2: UDINT;                 // 回路 2 模式切换审计计数 [次] / Loop 2 switch audit count
    uErrCode  : UDINT;                 // 信息级码，0 = 无信息 / Info-level code, 0 = none
    bValid    : BOOL;                  // 输出可用标志 / Outputs usable flag
END_VAR
VAR
    trigAuto1 : R_TRIG;                // 回路 1 自动请求沿，每拍无条件刷新 / Loop 1 auto edge, refreshed every scan
    trigMan1  : R_TRIG;                // 回路 1 手动请求沿，每拍无条件刷新 / Loop 1 manual edge, refreshed every scan
    trigAuto2 : R_TRIG;                // 回路 2 自动请求沿，每拍无条件刷新 / Loop 2 auto edge, refreshed every scan
    trigMan2  : R_TRIG;                // 回路 2 手动请求沿，每拍无条件刷新 / Loop 2 manual edge, refreshed every scan
    _bSw1     : BOOL;                  // 回路 1 切换脉冲内部暂存（统一出口映射） / Loop 1 switch stage
    _bSw2     : BOOL;                  // 回路 2 切换脉冲内部暂存（统一出口映射） / Loop 2 switch stage
END_VAR
VAR CONSTANT
    DL_HA_AUDIT_MAX  : UDINT := 4294967295; // 审计计数上限（饱和不回绕）/ Audit count ceiling, saturating
    DL_HA_CODE_KEY1  : UDINT := 16#0005_3060; // 信息级：回路 1 单钥匙拒绝码 / Info code: loop 1 single key refused
    DL_HA_CODE_KEY2  : UDINT := 16#0005_3061; // 信息级：回路 2 单钥匙拒绝码 / Info code: loop 2 single key refused
    DL_HA_CODE_SAT   : UDINT := 16#0005_3062; // 信息级：审计计数饱和码 / Info code: audit count saturated
END_VAR

// ---- 段 1｜沿实例无条件刷新 + 单拍脉冲出口预清（红线 R7 + 两段式）----
trigAuto1(CLK := bAutoReq1);          // 回路 1 自动沿每拍刷新 / Loop 1 auto edge refreshed
trigMan1(CLK := bManReq1);            // 回路 1 手动沿每拍刷新 / Loop 1 manual edge refreshed
trigAuto2(CLK := bAutoReq2);          // 回路 2 自动沿每拍刷新 / Loop 2 auto edge refreshed
trigMan2(CLK := bManReq2);            // 回路 2 手动沿每拍刷新 / Loop 2 manual edge refreshed
_bSw1 := FALSE;                       // 回路 1 切换暂存先清零 / Loop 1 switch stage cleared
_bSw2 := FALSE;                       // 回路 2 切换暂存先清零 / Loop 2 switch stage cleared
uErrCode := 16#0000_0000;             // 信息码每拍重算（信息级不锁存）/ Info code recomputed, never latched

// ---- 段 2｜回路 1 模式状态机（CASE 带 ELSE；双钥匙闸前置）----
CASE eMode1 OF
    E_DL_HaMode.eAuto:                 // 自动相：可切手动（双钥匙闸）
        IF trigMan1.Q THEN             // 手动请求沿
            IF bKeyA1 AND bKeyB1 THEN  // 双钥匙确认闸 / Dual-key gate
                eMode1 := E_DL_HaMode.eManual; // 切手动 / To manual
                _bSw1 := TRUE;         // 切换脉冲内部置位（出口统一映射）/ Switch stage set
                IF uAuditCnt1 < DL_HA_AUDIT_MAX THEN
                    uAuditCnt1 := uAuditCnt1 + 1; // 审计计数推进 / Audit count advance
                ELSE
                    uErrCode := DL_HA_CODE_SAT;   // 审计计数饱和留痕 / Audit saturation trace
                END_IF
            ELSE
                uErrCode := DL_HA_CODE_KEY1; // 单钥匙拒绝留痕（不切换）/ Single-key refusal, no switch
            END_IF
        END_IF
    E_DL_HaMode.eManual:               // 手动相：可切自动（双钥匙闸）
        IF trigAuto1.Q THEN            // 自动请求沿
            IF bKeyA1 AND bKeyB1 THEN  // 双钥匙确认闸 / Dual-key gate
                eMode1 := E_DL_HaMode.eAuto;   // 切自动 / To auto
                _bSw1 := TRUE;         // 切换脉冲内部置位 / Switch stage set
                IF uAuditCnt1 < DL_HA_AUDIT_MAX THEN
                    uAuditCnt1 := uAuditCnt1 + 1; // 审计计数推进 / Audit count advance
                ELSE
                    uErrCode := DL_HA_CODE_SAT;   // 审计计数饱和留痕 / Audit saturation trace
                END_IF
            ELSE
                uErrCode := DL_HA_CODE_KEY1; // 单钥匙拒绝留痕（不切换）/ Single-key refusal, no switch
            END_IF
        END_IF
    ELSE                               // 非法模式兜底（R21：CASE 必带 ELSE）
        eMode1 := E_DL_HaMode.eManual; // 拦截非法值归手动（人工介入侧安全）/ Catch illegal value to manual, safe side
END_CASE

// ---- 段 3｜回路 2 模式状态机（同段 2 口径）----
CASE eMode2 OF
    E_DL_HaMode.eAuto:                 // 自动相：可切手动（双钥匙闸）
        IF trigMan2.Q THEN             // 手动请求沿
            IF bKeyA2 AND bKeyB2 THEN  // 双钥匙确认闸 / Dual-key gate
                eMode2 := E_DL_HaMode.eManual; // 切手动 / To manual
                _bSw2 := TRUE;         // 切换脉冲内部置位 / Switch stage set
                IF uAuditCnt2 < DL_HA_AUDIT_MAX THEN
                    uAuditCnt2 := uAuditCnt2 + 1; // 审计计数推进 / Audit count advance
                ELSE
                    uErrCode := DL_HA_CODE_SAT;   // 审计计数饱和留痕 / Audit saturation trace
                END_IF
            ELSE
                uErrCode := DL_HA_CODE_KEY2; // 单钥匙拒绝留痕（不切换）/ Single-key refusal, no switch
            END_IF
        END_IF
    E_DL_HaMode.eManual:               // 手动相：可切自动（双钥匙闸）
        IF trigAuto2.Q THEN            // 自动请求沿
            IF bKeyA2 AND bKeyB2 THEN  // 双钥匙确认闸 / Dual-key gate
                eMode2 := E_DL_HaMode.eAuto;   // 切自动 / To auto
                _bSw2 := TRUE;         // 切换脉冲内部置位 / Switch stage set
                IF uAuditCnt2 < DL_HA_AUDIT_MAX THEN
                    uAuditCnt2 := uAuditCnt2 + 1; // 审计计数推进 / Audit count advance
                ELSE
                    uErrCode := DL_HA_CODE_SAT;   // 审计计数饱和留痕 / Audit saturation trace
                END_IF
            ELSE
                uErrCode := DL_HA_CODE_KEY2; // 单钥匙拒绝留痕（不切换）/ Single-key refusal, no switch
            END_IF
        END_IF
    ELSE                               // 非法模式兜底（R21：CASE 必带 ELSE）
        eMode2 := E_DL_HaMode.eManual; // 拦截非法值归手动 / Catch illegal value to manual
END_CASE

// ---- 段 4｜统一出口：切换脉冲单拍映射（两段式）----
bSwitchPulse1 := _bSw1;               // 回路 1 切换脉冲本拍有效 / Loop 1 pulse valid this scan
bSwitchPulse2 := _bSw2;               // 回路 2 切换脉冲本拍有效 / Loop 2 pulse valid this scan
bValid := TRUE;                       // 输出恒可用 / Outputs always usable
END_FUNCTION_BLOCK

(* ---- FB_DL_HeadboxJetRatioLoop.st ---- *)
(*
  DL Factory R84 | FB_DL_HeadboxJetRatioLoop
  功能：流浆箱唇口喷射比闭环：由浆料流量、浆浓、幅宽与唇口开度换算浆速并求喷射比，按喷射比偏差与五点横幅定量偏差加权均值出 PI 唇口开度指令，限位时冻结积分并出限位位，网速或开度为零时不出比值保持上一有效指令。
  开源溯源：无（clean-room 自研，依据公开工艺公式与安全设计惯例，来源=行业通用公式+工程实践，许可证=MIT，借鉴点=公式结构与联锁分层）
  规则：R1-R16 全遵守
  ------------------------------------------------------------------
  分类 DL_Process ｜ 复杂度 cx4 ｜ 版本 v1.0.0 ｜ 平台 纯 IEC 61131-3（TON、R_TRIG、LREAL、ENUM、CASE）
  边界一：只出唇口开度指令与限位位，不驱动唇口伺服、不控上浆泵、不改横幅执行器（属主边界，执行由下层 PRG 完成）。
  边界二：浆速换算——浆速 [m/min]＝浆料流量 [L/min] ÷（唇口开度 [mm] × 幅宽 [m]），
          推导：流量 [L/min]＝0.001 [m³/L] × 数值，面积 [m²]＝0.001 [m/mm] × 开度 × 幅宽，
          两者相除后两个 0.001 相消，故公式不含任何折算系数（量纲自洽，写死为字面量形式）。
  边界三：喷射比＝浆速 ÷ 网速，为使浆速与网速同速，目标喷射比 fJetRatioSp 默认 1.00（唇口射流与网速等速为常规稳态）。
  边界四：横幅定量偏差五点加权——权重为三角权 1／2／3／2／1（中心权重三、两侧递减），权数和为常量 9；
          权重按 3 − ABS(i − 2) 逐点算术生成，不建常量权重表（避免定长数组常量在部分平台不被接受）。
  边界五：控制律为位置式 PI——开度指令＝基准开度 ＋ Kp·e ＋ 积分项，积分项在限位或相位不在调节窗口时冻结（抗饱和）；
          基准开度在进入稳定相时锁存为当时的开度指令（复位与首扫时该指令以开度反馈为初值），故积分项归零时指令自然回到基准，无扰切换。
  边界六：无效拍语义——网速或当前开度为零（或非有限）→ 不计算喷射比、xValid 出假、开度指令保持上一有效值，
          相位与积分均不推进（不除零、不外推）。
  量纲自检：喷射比 [-]＝浆速 [m/min] ÷ 网速 [m/min]；开度 [mm]＝fSliceMm、fSliceCmd、上下限；
          流量 [L/min]＝fStockFlowLpm；浓度 [百分数]＝fConsPct 与 fConsNomPct；幅宽 [m]＝fWidthM；
          横幅偏差 [g/m²]＝afProfileDev 五点；增益 Kp 单位 [mm/比值]、Ki 单位 [mm/比值·拍]。
  码表：本件全部码位为信息级（2901 组态越域、2902 入参非有限、2903 网速或开度为零、2904 开度到达限位、
        2905 非法相位）；信息级码每拍重算且不置 bError；限位由 xAtLimit 电平位表达，故本件无 bError 出口（R187）。
  输出契约：fSliceCmd 在上下限之间恒成立（域内硬钳）；xAtLimit 为电平位（限位相成立期间为真）；
          fJetRatio 在无有效比值的拍保持上一有效值；fProfileMean 为五点加权横幅偏差 [g/m²]。
  修订记录：2026-11-24 v1.0.0 R84 首版（批 R84 · 序号 44）
*)

TYPE E_DL_HjrState :
(
    eIdle      := 0, // 空闲：等使能与输入有效 / idle, waiting for the enable and valid inputs
    eStabilize := 10, // 稳定：等稳定窗到期或偏差入死区 / stabilising, waiting for the window or the dead band
    eRegulate  := 20, // 调节：闭环出开度指令 / regulating, the loop drives the slice
    eLimitHold := 30  // 限位保持：开度到限，冻结积分 / limit hold, the slice is on a limit and the integral is frozen
);
END_TYPE

TYPE E_DL_HjrCause :
(
    eNone      := 0, // 无成因 / no cause
    eCfgBad    := 1, // 组态越域（信息级 2901）/ the configuration is out of domain, info grade 2901
    eNotFinite := 2, // 入参非有限（信息级 2902）/ a non-finite input, info grade 2902
    eNoRatio   := 3, // 网速或开度为零（信息级 2903）/ the wire speed or the slice is zero, info grade 2903
    eAtLimit   := 4, // 开度到达限位（信息级 2904）/ the slice reached a limit, info grade 2904
    ePhaseBad  := 5  // 非法相位（信息级 2905）/ an illegal phase, info grade 2905
);
END_TYPE

FUNCTION_BLOCK FB_DL_HeadboxJetRatioLoop
VAR CONSTANT
    DL_HJR_KP          : LREAL := 0.30;    // 比例增益 [mm/比值] / the proportional gain [mm per ratio]
    DL_HJR_KI          : LREAL := 0.02;    // 积分增益（每拍）[mm/比值·拍] / the integral gain per scan [mm per ratio]
    DL_HJR_INT_MAX     : LREAL := 0.60;    // 积分项限幅 [mm] / the integral term limit [mm]
    DL_HJR_STEP_MM     : LREAL := 0.05;    // 单拍开度变化限幅 [mm] / the per scan slice step limit [mm]
    DL_HJR_DEADBAND    : LREAL := 0.01;    // 喷射比死区 [比值] / the jet ratio dead band [ratio]
    DL_HJR_PROF_GAIN   : LREAL := 0.05;    // 横幅偏差折算增益 [比值/(g/m²)] / the profile deviation gain [ratio per g/m2]
    DL_HJR_CONS_GAIN   : LREAL := 0.50;    // 浆浓前馈增益 [mm/倍] / the consistency feed forward gain [mm per times]
    DL_HJR_LIMIT_BAND  : LREAL := 0.001;   // 限位判定带 [mm] / the limit detection band [mm]
    DL_HJR_W_CENTER    : INT := 3;         // 横幅权重基数（中心权重）[-] / the centre weight of the profile weights [-]
    DL_HJR_W_LAST      : INT := 4;         // 横幅最后一点下标 [-] / the last profile subscript [-]
    DL_HJR_EPS         : LREAL := 1.0E-9;  // 除法零闸与零判定门限 [-] / the division guard and zero test threshold [-]
END_VAR
VAR_INPUT
    bEnable        : BOOL := TRUE;      // 使能，失能回空闲且冻结积分 [-] / enable, a disable returns to idle and freezes the integral
    bReset         : BOOL := FALSE;     // 复位上升沿清积分与基准开度 [-] / reset rising edge clears the integral and the base
    fStockFlowLpm  : LREAL := 6000.0;   // 浆料流量 [L/min] / the stock flow [L/min]
    fConsPct       : LREAL := 3.20;     // 浆浓（实测）[百分数] / the measured consistency [percent]
    fConsNomPct    : LREAL := 3.20;     // 浆浓设计值（前馈基准）[百分数] / the design consistency as the feed forward base [percent]
    fWireSpeedMpm  : LREAL := 800.0;    // 网速 [m/min] / the wire speed [m/min]
    fSliceMm       : LREAL := 9.00;     // 唇口开度反馈 [mm] / the slice opening feedback [mm]
    fSliceMinMm    : LREAL := 3.00;     // 唇口开度下限 [mm] / the slice lower limit [mm]
    fSliceMaxMm    : LREAL := 20.0;     // 唇口开度上限 [mm] / the slice upper limit [mm]
    fWidthM        : LREAL := 6.00;     // 成形幅宽 [m] / the forming width [m]
    fJetRatioSp    : LREAL := 1.00;     // 目标喷射比（默认等速）[比值] / the jet ratio setpoint, unity by default [ratio]
    afProfileDev   : ARRAY[0..4] OF LREAL := [0.0, 0.0, 0.0, 0.0, 0.0]; // 横幅五点定量偏差 [g/m²] / the five point basis weight deviations [g/m2]
    tStab          : TIME := T#10S;     // 稳定窗（进稳定相后计时）[毫秒] / the stabilising window [ms]
END_VAR
VAR_OUTPUT
    fSliceCmd      : LREAL := 0.0;  // 唇口开度指令 [mm] / the slice opening command [mm]
    fJetRatio      : LREAL := 1.0;  // 实测喷射比（无有效值时保持）[比值] / the measured jet ratio, held when invalid [ratio]
    fStockSpeedMpm : LREAL := 0.0;  // 换算浆速 [m/min] / the converted stock speed [m/min]
    fProfileMean   : LREAL := 0.0;  // 横幅五点加权偏差均值 [g/m²] / the weighted profile deviation mean [g/m2]
    fRatioErr      : LREAL := 0.0;  // 喷射比偏差（含前馈与横幅修正）[比值] / the ratio error including both corrections [ratio]
    fSliceStep     : LREAL := 0.0;  // 本拍开度增量（限幅后）[mm] / the slice step of this scan after limiting [mm]
    xAtLimit       : BOOL := FALSE; // 开度到达限位（电平位）[-] / the slice reached a limit
    eState         : E_DL_HjrState := E_DL_HjrState.eIdle; // 相位出口 [枚举] / the phase outlet [enum]
    iErrCode       : INT := 0;      // 信息级码（每拍重算，非锁存）[码] / the info grade code, recomputed every scan [code]
    xValid         : BOOL := FALSE; // 本拍输入可信且比值可算 [-] / the inputs are trustworthy and the ratio is computable
END_VAR
VAR
    rtReset    : R_TRIG; // 复位沿实例（无量纲）[-] / the reset edge refreshed unconditionally
    tonStab    : TON;    // 稳定窗实例（无量纲）[-] / the stabilising window gated by eStabilize
    _eState    : E_DL_HjrState := E_DL_HjrState.eIdle; // 内部相位（枚举，无量纲）[-] / the internal phase, the only CASE target
    _i         : INT := 0;      // 横幅遍历下标 [-] / the profile traversal index
    _iErrTmp   : INT := 0;      // 本拍信息级码暂存 [码] / the scan info code scratch [code]
    _bInit     : BOOL := FALSE; // 首扫初始化完成标志（R310）[-] / the first scan initialisation flag
    _bScalarFin: BOOL := FALSE; // 标量浮点入参有限 [-] / the scalar floating inputs are finite
    _bProfFin  : BOOL := FALSE; // 横幅五点数组逐点有限 [-] / every profile point is finite
    _bFinOk    : BOOL := FALSE; // 标量与数组有限之合取 [-] / the conjunction of the scalar and array gates
    _bCfgOk    : BOOL := FALSE; // 组态参数域内 [-] / the configuration is inside its domain
    _bRatioOk  : BOOL := FALSE; // 网速与开度非零（比值可算）[-] / the wire speed and the slice are non zero
    _bAtLimit  : BOOL := FALSE; // 开度到达限位判据 [-] / the slice limit verdict
    _bFreeze   : BOOL := FALSE; // 积分冻结判据 [-] / the integral freeze verdict
    _fStockVel : LREAL := 0.0;  // 换算浆速（本拍）[m/min] / the converted stock speed of this scan [m/min]
    _fRatio    : LREAL := 1.0;  // 喷射比（本拍计算）[比值] / the jet ratio of this scan [ratio]
    _fRatioLst : LREAL := 1.0;  // 上一有效喷射比（保持槽）[比值] / the last valid jet ratio, a hold slot [ratio]
    _fWSum     : LREAL := 0.0;  // 横幅权重和 [-] / the sum of the profile weights
    _fDevSum   : LREAL := 0.0;  // 横幅加权偏差和 [g/m²] / the weighted profile deviation sum [g/m2]
    _fW        : LREAL := 0.0;  // 单点权重 [-] / the single point weight
    _fProfMean : LREAL := 0.0;  // 横幅加权均值 [g/m²] / the weighted profile mean [g/m2]
    _fConsFact : LREAL := 1.0;  // 浆浓与设计值之比（前馈）[倍] / the consistency ratio for the feed forward [times]
    _fErr      : LREAL := 0.0;  // 喷射比偏差（原始）[比值] / the raw ratio error [ratio]
    _fErrCtl   : LREAL := 0.0;  // 加前馈与横幅修正后的控制偏差 [比值] / the control error with both corrections [ratio]
    _fInt      : LREAL := 0.0;  // 积分项（位置式，限幅）[mm] / the integral term of the positional form [mm]
    _fBase     : LREAL := 0.0;  // 基准开度（进稳定相时锁存）[mm] / the base opening latched when stabilising starts [mm]
    _fPiOut    : LREAL := 0.0;  // PI 输出量 [mm] / the PI output [mm]
    _fTarget   : LREAL := 0.0;  // 目标开度（未限幅）[mm] / the target opening before limiting [mm]
    _fStep     : LREAL := 0.0;  // 本拍开度增量（限幅后）[mm] / the step of this scan after limiting [mm]
    _fCmd      : LREAL := 0.0;  // 开度指令累加（唯一写入点）[mm] / the command accumulator, the only write point [mm]
    _fCmdLst   : LREAL := 0.0;  // 上一有效开度指令（无效拍保持）[mm] / the last valid command held on an invalid scan [mm]
    _tStab     : TIME := T#1S;  // 稳定窗实参（钳定后）[毫秒] / the stabilising window passed to the timer [ms]
END_VAR
// 段 0｜出口预置：全部出口先赋安全侧值，任何路径不留未初始化输出
xValid := FALSE; // 有效性预置假 / validity preset false
xAtLimit := FALSE; // 限位位预置假 / the limit bit preset false
fSliceCmd := _fCmdLst; // 开度指令回放上一有效值（无效拍保持，边界六）/ replay the last valid command
fJetRatio := _fRatioLst; // 喷射比回放上一有效值 / replay the last valid ratio
fStockSpeedMpm := 0.0; // 浆速预置零 / the stock speed preset zero
fProfileMean := 0.0; // 横幅均值预置零 / the profile mean preset zero
fRatioErr := 0.0; // 偏差预置零 / the error preset zero
fSliceStep := 0.0; // 开度增量预置零（不调节拍不出量）/ the step preset zero
eState := _eState; // 相位回放 / replay the phase
iErrCode := 0; // 信息级码预置零（本拍重算）/ the info code preset zero
_iErrTmp := 0; // 单拍码暂存预清（FB32-1）/ preclear the code scratch
_fStep := 0.0; // 单拍增量预清 / preclear the step
// 段 1｜非有限闸（标量）：NaN 自反比较、Inf 差值自减双判，逐项枚举九个标量浮点入参（R79、R272）
_bScalarFin := (fStockFlowLpm = fStockFlowLpm) AND ((fStockFlowLpm - fStockFlowLpm) = (fStockFlowLpm - fStockFlowLpm)) // 浆料流量有限 [-] / the stock flow is finite
    AND (fConsPct = fConsPct) AND ((fConsPct - fConsPct) = (fConsPct - fConsPct)) // 浆浓有限 [-] / the consistency is finite
    AND (fConsNomPct = fConsNomPct) AND ((fConsNomPct - fConsNomPct) = (fConsNomPct - fConsNomPct)) // 设计浆浓有限 [-] / the design consistency is finite
    AND (fWireSpeedMpm = fWireSpeedMpm) AND ((fWireSpeedMpm - fWireSpeedMpm) = (fWireSpeedMpm - fWireSpeedMpm)) // 网速有限 [-] / the wire speed is finite
    AND (fSliceMm = fSliceMm) AND ((fSliceMm - fSliceMm) = (fSliceMm - fSliceMm)) // 开度反馈有限 [-] / the slice feedback is finite
    AND (fSliceMinMm = fSliceMinMm) AND ((fSliceMinMm - fSliceMinMm) = (fSliceMinMm - fSliceMinMm)) // 开度下限有限 [-] / the slice floor is finite
    AND (fSliceMaxMm = fSliceMaxMm) AND ((fSliceMaxMm - fSliceMaxMm) = (fSliceMaxMm - fSliceMaxMm)) // 开度上限有限 [-] / the slice ceiling is finite
    AND (fWidthM = fWidthM) AND ((fWidthM - fWidthM) = (fWidthM - fWidthM)) // 幅宽有限 [-] / the width is finite
    AND (fJetRatioSp = fJetRatioSp) AND ((fJetRatioSp - fJetRatioSp) = (fJetRatioSp - fJetRatioSp)); // 目标喷射比有限 [-] / the setpoint is finite
// 段 2｜非有限闸（横幅数组）：逐点枚举，漏判单点会污染加权均值（R151）
_bProfFin := TRUE; // 逐点闸初值真 / the per point gate starts true
FOR _i := 0 TO (DL_HJR_W_LAST) DO // 定长字面界 0..4（禁动态上下界，E037）/ the literal subscript range
    IF NOT (afProfileDev[_i] = afProfileDev[_i]) THEN _bProfFin := FALSE; END_IF // 该点 NaN 判否 / the point is NaN
    IF (afProfileDev[_i] - afProfileDev[_i]) <> (afProfileDev[_i] - afProfileDev[_i]) THEN _bProfFin := FALSE; END_IF // 该点 Inf 判否 / the point is infinite
END_FOR
_bFinOk := _bScalarFin AND _bProfFin; // 标量与数组有限之合取 / the conjunction of the scalar and array gates
// 段 3｜组态域闸：开度上下限次序、幅宽与设计浆浓正定、稳定窗正定（R151）
_bCfgOk := (fSliceMinMm > 0.0) AND (fSliceMaxMm > fSliceMinMm) // 开度域闸（上限严格大于下限）[-] / the slice domain gate
    AND (fWidthM > DL_HJR_EPS) AND (fConsNomPct > DL_HJR_EPS) // 幅宽与设计浆浓非零 [-] / the width and the design consistency are non zero
    AND (fJetRatioSp > DL_HJR_EPS) AND (tStab > T#0S); // 目标比值与稳定窗域闸 [-] / the setpoint and the window gates
_tStab := tStab; // 稳定窗一级回退：取引脚值 [ms] / level one fallback, take the pin value
IF _tStab <= T#0S THEN _tStab := T#1S; END_IF // 稳定窗二级回退：按有效域钳定 / level two, clamp into the valid domain
IF NOT _bFinOk THEN _iErrTmp := 2902; ELSIF NOT _bCfgOk THEN _iErrTmp := 2901; END_IF // 信息级码分派（有限 → 组态）/ the info code dispatch
// 段 4｜首扫初始化与复位沿同块，作用域逐项声明（R310、R311）
IF (NOT _bInit) OR rtReset.Q THEN // 首扫一拍或复位沿 / the first scan or the reset edge
    _bInit := TRUE; // 首扫完成标志 / the first scan flag
    _fInt := 0.0; // 作用域一：清积分项（唯一清除边，R188）/ scope one, clear the integral term
    _fCmd := fSliceMm; // 作用域二：指令基准取当前反馈 [mm] / scope two, the command base is the feedback [mm]
    IF _fCmd < fSliceMinMm THEN _fCmd := fSliceMinMm; END_IF // 基准下限钳定 / clamp the base low
    IF _fCmd > fSliceMaxMm THEN _fCmd := fSliceMaxMm; END_IF // 基准上限钳定 / clamp the base high
    _fCmdLst := _fCmd; // 作用域二：上一有效指令同步 / scope two, sync the last valid command
    _fBase := _fCmd; // 作用域二：基准开度同步 / scope two, sync the base opening
    _fRatioLst := fJetRatioSp; // 作用域三：喷射比保持槽预置为目标值 / scope three, preset the ratio hold slot
    _eState := E_DL_HjrState.eIdle; // 作用域一：迁回空闲相 / scope one, migrate to idle
END_IF
// 段 5｜定时器与沿检测无条件周期刷新（R7），稳定窗只串 eStabilize 相
rtReset(CLK := bReset); // 复位沿无条件刷新 / unconditional refresh of the reset edge
tonStab(IN := (_eState = E_DL_HjrState.eStabilize) AND _bFinOk, PT := _tStab); // 稳定窗，只串稳定相 / the window gated by the stabilise phase
// 段 6｜横幅五点加权均值：三角权 1/2/3/2/1，权数和为常量九，除零结构性排除
_fWSum := 0.0; _fDevSum := 0.0; // 权重和与加权和清零 / clear the weight sum and the weighted sum
FOR _i := 0 TO (DL_HJR_W_LAST) DO // 定长字面界 0..4 / the literal subscript range
    _fW := INT_TO_LREAL(DL_HJR_W_CENTER - ABS(_i - 2)); // 三角权重 1/2/3/2/1 [-] / the triangular weight
    _fWSum := _fWSum + _fW; // 权重累加 / accumulate the weight
    _fDevSum := _fDevSum + (_fW * afProfileDev[_i]); // 加权偏差累加 [g/m²] / accumulate the weighted deviation
END_FOR
IF _fWSum > DL_HJR_EPS THEN // 权重和零闸（常量九，结构性恒真，防御性保留）/ the weight sum guard
    _fProfMean := _fDevSum / _fWSum; // 加权均值 [g/m²] / the weighted mean [g/m2]
ELSE // 权重和非法 / an illegal weight sum
    _fProfMean := 0.0; // 均值出零（不放大修正）/ the mean goes to zero
END_IF
IF NOT (_fProfMean = _fProfMean) THEN _fProfMean := 0.0; END_IF // 均值 NaN 兜底 / the NaN fallback
IF (_fProfMean - _fProfMean) <> (_fProfMean - _fProfMean) THEN _fProfMean := 0.0; END_IF // 均值 Inf 兜底 / the Inf fallback
// 段 7｜浆速与喷射比：网速或开度为零不计算比值，保持上一有效值（边界六、R4）
_bRatioOk := (ABS(fWireSpeedMpm) > DL_HJR_EPS) AND (ABS(fSliceMm) > DL_HJR_EPS) AND (ABS(fWidthM) > DL_HJR_EPS); // 三分母零闸 / the three denominator guards
IF _bRatioOk AND _bFinOk THEN // 比值可算且入参可信 / the ratio is computable with trustworthy inputs
    _fStockVel := fStockFlowLpm / (fSliceMm * fWidthM); // 浆速 [m/min]（两个千分折算相消，边界二）/ the stock speed [m/min]
    _fRatio := _fStockVel / fWireSpeedMpm; // 喷射比 [比值] / the jet ratio [ratio]
    IF NOT (_fRatio = _fRatio) THEN _fRatio := _fRatioLst; END_IF // 比值 NaN 兜底（回退上一有效）/ the NaN fallback to the hold slot
    IF (_fRatio - _fRatio) <> (_fRatio - _fRatio) THEN _fRatio := _fRatioLst; END_IF // 比值 Inf 兜底 / the Inf fallback to the hold slot
    _fRatioLst := _fRatio; // 保持槽写入（已过非有限闸，R133）/ the guarded write into the hold slot
ELSE // 网速或开度为零 / the wire speed or the slice is zero
    _fRatio := _fRatioLst; // 比值保持上一有效值 / hold the last valid ratio
    _fStockVel := 0.0; // 浆速出零（不虚报）/ the stock speed goes to zero
    IF _iErrTmp = 0 THEN _iErrTmp := 2903; END_IF // 信息级：比值不可算 / the info code for an uncomputable ratio
END_IF
// 段 8｜PI 调节与限位抗饱和：仅在调节窗口内积分（状态量门控，R99）
_fConsFact := 1.0; // 浆浓比预置一 / the consistency ratio preset unity
IF fConsNomPct > DL_HJR_EPS THEN _fConsFact := fConsPct / fConsNomPct; END_IF // 浆浓比（分母已过域闸）[倍] / the consistency ratio [times]
IF _bRatioOk AND _bFinOk AND _bCfgOk AND bEnable THEN // 控制律在输入可信、比值可算且使能时推进（R583 补使能门控）
    _fErr := _fRatio - fJetRatioSp; // 喷射比偏差 [比值]，正为浆速偏高 / the ratio error, positive means a fast jet
    _fErrCtl := _fErr + (DL_HJR_PROF_GAIN * _fProfMean) + (DL_HJR_CONS_GAIN * (_fConsFact - 1.0)); // 加横幅修正与浆浓前馈 / add the profile and consistency corrections
    IF ABS(_fErrCtl) <= DL_HJR_DEADBAND THEN _fErrCtl := 0.0; END_IF // 死区内偏差取零（不踢动）/ zero the error inside the dead band
    _bFreeze := (_bAtLimit OR (_eState = E_DL_HjrState.eIdle) OR (_eState = E_DL_HjrState.eStabilize) OR (_eState = E_DL_HjrState.eLimitHold)) OR (NOT bEnable); // R583 补 eStabilize：稳定窗内不得积分，否则开窗期已积出超调 // 冻结判据挂状态量（R99）；限位为跨拍电平量，本处取上一拍限位态，限位持续期内每拍皆冻结，单拍滞后不影响抗饱和 / the freeze verdict uses the state, the limit is a level lasting many scans
    IF NOT _bFreeze THEN // 未冻结才积分 / integrate only while unfrozen
        _fInt := _fInt + (DL_HJR_KI * _fErrCtl); // 积分项累加 [mm] / accumulate the integral [mm]
        IF _fInt > DL_HJR_INT_MAX THEN _fInt := DL_HJR_INT_MAX; ELSIF _fInt < (0.0 - DL_HJR_INT_MAX) THEN _fInt := (0.0 - DL_HJR_INT_MAX); END_IF // 积分项双向限幅 / the integral limit
    END_IF
    _fPiOut := (DL_HJR_KP * _fErrCtl) + _fInt; // PI 输出 [mm] / the PI output [mm]
    _fTarget := _fBase + _fPiOut; // 目标开度 [mm] / the target opening [mm]
    _fStep := _fTarget - _fCmd; // 本拍应走增量 [mm] / the step required this scan [mm]
    IF _fStep > DL_HJR_STEP_MM THEN _fStep := DL_HJR_STEP_MM; ELSIF _fStep < (0.0 - DL_HJR_STEP_MM) THEN _fStep := (0.0 - DL_HJR_STEP_MM); END_IF // 单拍双向限幅 / the two sided step limit
    IF NOT (_fStep = _fStep) THEN _fStep := 0.0; END_IF // 增量 NaN 兜底 / the NaN fallback
    IF (_fStep - _fStep) <> (_fStep - _fStep) THEN _fStep := 0.0; END_IF // 增量 Inf 兜底 / the Inf fallback
    _fCmd := _fCmd + _fStep; // 指令累加（唯一写入点）[mm] / the only write point of the command [mm]
    IF _fCmd > fSliceMaxMm THEN _fCmd := fSliceMaxMm; END_IF // 上限硬钳 / the hard clamp high
    IF _fCmd < fSliceMinMm THEN _fCmd := fSliceMinMm; END_IF // 下限硬钳 / the hard clamp low
    _fCmdLst := _fCmd; // 上一有效指令同步 / sync the last valid command
END_IF
_bAtLimit := (_fCmd >= (fSliceMaxMm - DL_HJR_LIMIT_BAND)) OR (_fCmd <= (fSliceMinMm + DL_HJR_LIMIT_BAND)); // 限位判据（含判定带）/ the limit verdict with its band
// 段 9｜相位状态机：ENUM ＋ CASE ＋ ELSE 非法相位兜底（R6、R128）
CASE _eState OF
E_DL_HjrState.eIdle: // 空闲相：退出条件三（失能驻留、输入不可信驻留、使能且可信进取）
    IF bEnable AND _bFinOk AND _bCfgOk THEN // 使能且双闸通过 / enabled with both gates passed
        _fBase := _fCmd; // 基准开度锁存为当前指令 [mm] / latch the base opening [mm]
        _fInt := 0.0; // 积分项无扰归零（进稳定相）/ clear the integral on entry
        _eState := E_DL_HjrState.eStabilize; // 迁稳定相 / migrate to stabilise
    END_IF
E_DL_HjrState.eStabilize: // 稳定相：退出条件四（失能、限位、稳定窗到期、偏差入死区）
    IF NOT bEnable THEN // 使能丢失 / the enable was lost
        _eState := E_DL_HjrState.eIdle; // 回空闲 / back to idle
    ELSIF _bAtLimit THEN // 一进入即到限 / already on a limit
        _eState := E_DL_HjrState.eLimitHold; // 迁限位相 / migrate to the limit hold
    ELSIF tonStab.Q THEN // 稳定窗到期 / the window expired
        _eState := E_DL_HjrState.eRegulate; // 迁调节相 / migrate to regulate
    ELSIF ABS(_fErrCtl) <= DL_HJR_DEADBAND THEN // 偏差已入死区（无需调节）/ the error already sits in the dead band
        _eState := E_DL_HjrState.eRegulate; // 迁调节相（保持指令）/ migrate to regulate
    END_IF
E_DL_HjrState.eRegulate: // 调节相：退出条件三（失能、限位、输入不可信）
    IF NOT bEnable THEN // 使能丢失 / the enable was lost
        _eState := E_DL_HjrState.eIdle; // 回空闲 / back to idle
    ELSIF _bAtLimit THEN // 开度到达限位 / the slice reached a limit
        _eState := E_DL_HjrState.eLimitHold; // 迁限位相（冻结积分）/ migrate to the limit hold
    ELSIF NOT _bFinOk THEN // 输入不可信（停在本相但不出量）/ the inputs are untrustworthy
        _eState := E_DL_HjrState.eIdle; // 回空闲等恢复 / back to idle
    END_IF
E_DL_HjrState.eLimitHold: // 限位相：退出条件二（失能、限位条件消失）
    IF NOT bEnable THEN // 使能丢失 / the enable was lost
        _eState := E_DL_HjrState.eIdle; // 回空闲 / back to idle
    ELSIF NOT _bAtLimit THEN // 限位条件消失 / the limit condition cleared
        _eState := E_DL_HjrState.eRegulate; // 回调节相 / back to regulate
    END_IF
ELSE // 非法相位兜底（R6、R128）
    _eState := E_DL_HjrState.eIdle; // 回安全态空闲 / back to the safe idle phase
    _iErrTmp := 2905; // 信息级非法相位码 / the info grade illegal phase code
END_CASE
IF _bAtLimit AND (_iErrTmp = 0) THEN _iErrTmp := 2904; END_IF // 限位信息级码（电平位另由 xAtLimit 表达）/ the limit info code
// 段 10｜统一出口：单点映射，限位位与指令同源（R191、FB51-3）
eState := _eState; // 相位单点映射 / the single point mapping of the phase
xAtLimit := _bAtLimit; // 限位位单点映射 / the single point mapping of the limit bit
fSliceCmd := _fCmdLst; // 开度指令单点映射（无效拍保持上一有效值，边界六）/ the command mapping with the hold
fJetRatio := _fRatioLst; // 喷射比单点映射（无效拍保持上一有效值）/ the ratio mapping with the hold
fStockSpeedMpm := _fStockVel; // 浆速单点映射 [m/min] / the stock speed mapping [m/min]
fProfileMean := _fProfMean; // 横幅均值单点映射 [g/m²] / the profile mean mapping [g/m2]
fRatioErr := _fErrCtl; // 控制偏差单点映射 [比值] / the control error mapping [ratio]
fSliceStep := _fStep; // 开度增量单点映射 [mm] / the step mapping [mm]
iErrCode := _iErrTmp; // 信息级码单点映射（每拍重算，不锁存）/ the info code mapping
xValid := _bFinOk AND _bCfgOk AND _bRatioOk AND (_iErrTmp <> 2905); // 有效性：三闸通过且非非法相位（限位码 2904 不影响有效性）/ valid unless the phase is illegal
END_FUNCTION_BLOCK

(* ---- FB_DL_HeadboxSliceSeq.st ---- *)
(*
  DL Factory R84 | FB_DL_HeadboxSliceSeq
  功能：流浆箱唇口开度调节时序，含开度限位、粗调/精调分级与调节死区
  开源溯源：无（clean-room 自研，依据公开工艺公式，来源=行业通用公式，许可证=MIT，借鉴点=公式结构）
  规则：R1-R16 全遵守
*)
TYPE E_DL_HbSliceState :
(
    eIdle := 0, // 空闲待命 [-] / idle [-]
    ePrePos := 1, // 粗定位相 [-] / coarse positioning phase [-]
    eFineAdj := 2, // 精调相 [-] / fine adjustment phase [-]
    eStableCheck := 3, // 稳定确认相 [-] / stability confirmation phase [-]
    eReady := 4, // 就绪相 [-] / ready phase [-]
    eFault := 5 // 故障锁存相 [-] / fault latched phase [-]
) := eIdle;
END_TYPE

FUNCTION_BLOCK FB_DL_HeadboxSliceSeq
VAR_INPUT
    xStart : BOOL; // 唇口调节启动命令 [-] / slice adjustment start command [-]
    xReset : BOOL; // 复位命令，上升沿清故障码 [-] / reset command [-]
    rSliceAct : REAL; // 唇口开度实测值 [mm] / measured slice opening [mm]
    rSliceTarget : REAL := 12.0; // 唇口目标开度 [mm] / target slice opening [mm]
    fPosMinMm : REAL := 5.0; // 开度机械下限 [mm] / mechanical lower limit [mm]
    fPosMaxMm : REAL := 25.0; // 开度机械上限 [mm] / mechanical upper limit [mm]
    fCoarseBandMm : REAL := 0.5; // 粗调转入精调的带宽 [mm] / coarse to fine handover band [mm]
    fDeadbandMm : REAL := 0.05; // 精调调节死区 [mm] / fine adjustment deadband [mm]
    fCoarseStepMm : REAL := 0.20; // 粗调每拍步长 [mm] / coarse step per scan [mm]
    fFineStepMm : REAL := 0.02; // 精调每拍步长 [mm] / fine step per scan [mm]
    tPreLimit : TIME := T#60S; // 粗定位超时 [s] / coarse positioning timeout [s]
    tFineLimit : TIME := T#30S; // 精调超时 [s] / fine adjustment timeout [s]
    tStableLimit : TIME := T#5S; // 稳定确认时长 [s] / stability confirmation duration [s]
END_VAR
VAR_OUTPUT
    eState : E_DL_HbSliceState; // 当前时序状态 [-] / current sequence state [-]
    rSlicePos : REAL; // 唇口开度指令（限位后） [mm] / slice opening command after limiting [mm]
    iErrCode : INT; // 故障码 0=正常，801~805 [-] / error code, 801 to 805 [code]
    xReady : BOOL; // 开度就绪 [-] / opening ready [-]
END_VAR
VAR
    rtStart : R_TRIG; // 启动上升沿实例 [-] / start rising edge instance [-]
    rtReset : R_TRIG; // 复位上升沿实例 [-] / reset edge instance [-]
    tonPre : TON; // 粗定位超时定时器 [-] / coarse positioning timer [-]
    tonFine : TON; // 精调超时定时器 [-] / fine adjustment timer [-]
    tonStable : TON; // 稳定确认定时器 [-] / stability timer [-]
    _eState : E_DL_HbSliceState := E_DL_HbSliceState.eIdle; // 内部相位（CASE 唯一写目标） [-] / internal phase [-]
    _iErr : INT; // 故障码内部锁存 [-] / latched error code [-]
    rPos : REAL; // 开度指令内部量 [mm] / internal opening command [mm]
    rErrMm : REAL; // 开度偏差（目标 − 实测） [mm] / opening error [mm]
    xCfgBad : BOOL; // 组态非法当拍标志 [-] / illegal configuration flag [-]
END_VAR

// 段 0｜边沿与定时器实例无条件周期刷新（R7）
rtStart(CLK := xStart); // 启动沿每拍必调 [-] / start edge every scan [-]
rtReset(CLK := xReset); // 复位沿每拍必调 [-] / reset edge every scan [-]
tonPre(IN := _eState = E_DL_HbSliceState.ePrePos, PT := tPreLimit); // 粗定位相闸 [-] / coarse phase gate [-]
tonFine(IN := _eState = E_DL_HbSliceState.eFineAdj, PT := tFineLimit); // 精调相闸 [-] / fine phase gate [-]
tonStable(IN := _eState = E_DL_HbSliceState.eStableCheck, PT := tStableLimit); // 稳定相闸 [-] / stability phase gate [-]

// 段 1｜组态闸与当拍偏差派生（限位区间/死区/步长必须有效）
xCfgBad := NOT (fPosMinMm < fPosMaxMm) OR NOT (fDeadbandMm > 1.0E-9) OR NOT (fCoarseStepMm > 1.0E-9) OR NOT (fFineStepMm > 1.0E-9); // 限位/死区/步长正域闸（防除零） [mm] / limit, deadband and step gate [mm]
xCfgBad := xCfgBad OR NOT (rSliceAct > -1.0E30 AND rSliceAct < 1.0E30) OR NOT (rSliceTarget > -1.0E30 AND rSliceTarget < 1.0E30); // 开度非有限闸 [-] / non finite opening gate [-]
xCfgBad := xCfgBad OR (rSliceTarget < fPosMinMm) OR (rSliceTarget > fPosMaxMm); // 目标越限闸：不得超出机械限位 [mm] / target outside the mechanical limits [mm]
IF xCfgBad THEN
    _iErr := 801; // 组态非法码 [-] / illegal configuration code [-]
    _eState := E_DL_HbSliceState.eFault; // 锁存迁故障相 [-] / latch into the fault phase [-]
END_IF
rErrMm := rSliceTarget - rSliceAct; // mm − mm = mm / [mm] minus [mm] = [mm]

// 段 2｜复位沿：清故障码与相位（R189）
IF rtReset.Q THEN
    _iErr := 0; // 清故障码 [-] / clear error code [-]
    _eState := E_DL_HbSliceState.eIdle; // 回空闲相 [-] / back to idle [-]
END_IF

// 段 3｜主状态机（合法事件优先于超时迁移，R275）
CASE _eState OF
    E_DL_HbSliceState.eIdle: // 空闲相：指令跟随实测，无扰起步 [-] / idle [-]
        rPos := rSliceAct; // mm 直取 [mm] / take the measurement [mm]
        IF rtStart.Q THEN
            _eState := E_DL_HbSliceState.ePrePos; // 启动沿进粗定位相 [-] / start edge enters coarse positioning [-]
        END_IF
    E_DL_HbSliceState.ePrePos: // 粗定位相：大步长逼近 [-] / coarse positioning [-]
        IF ABS(rErrMm) <= fCoarseBandMm THEN
            _eState := E_DL_HbSliceState.eFineAdj; // 进入粗调带转精调相 [-] / inside the band leads to fine adjustment [-]
        ELSIF tonPre.Q THEN
            _iErr := 802; _eState := E_DL_HbSliceState.eFault; // 粗定位超时（执行机构卡涩） [-] / coarse positioning timeout [-]
        ELSE
            IF rErrMm > 0.0 THEN
                rPos := rPos + fCoarseStepMm; // mm + mm = mm（正向步进） / [mm] + [mm] = [mm]
            ELSE
                rPos := rPos - fCoarseStepMm; // mm − mm = mm（反向步进） / [mm] - [mm] = [mm]
            END_IF
        END_IF
    E_DL_HbSliceState.eFineAdj: // 精调相：小步长收敛至死区 [-] / fine adjustment [-]
        IF ABS(rErrMm) <= fDeadbandMm THEN
            _eState := E_DL_HbSliceState.eStableCheck; // 进死区转稳定确认 [-] / inside the deadband leads to stability check [-]
        ELSIF tonFine.Q THEN
            _iErr := 803; _eState := E_DL_HbSliceState.eFault; // 精调超时（无法收敛） [-] / fine adjustment timeout [-]
        ELSE
            IF rErrMm > 0.0 THEN
                rPos := rPos + fFineStepMm; // mm + mm = mm / [mm] + [mm] = [mm]
            ELSE
                rPos := rPos - fFineStepMm; // mm − mm = mm / [mm] - [mm] = [mm]
            END_IF
        END_IF
    E_DL_HbSliceState.eStableCheck: // 稳定确认相：死区内持续保持 [-] / stability confirmation [-]
        IF ABS(rErrMm) > (2.0 * fDeadbandMm) THEN
            _iErr := 804; _eState := E_DL_HbSliceState.eFault; // 稳定期漂出死区两倍（执行机构打滑） [-] / drifted out of twice the deadband [-]
        ELSIF tonStable.Q THEN
            _eState := E_DL_HbSliceState.eReady; // 稳定时长满转就绪相 [-] / stability elapsed leads to ready [-]
        END_IF
    E_DL_HbSliceState.eReady: // 就绪相 [-] / ready [-]
        IF NOT xStart THEN
            _eState := E_DL_HbSliceState.eIdle; // 命令撤销回空闲 [-] / command released returns to idle [-]
        END_IF
    E_DL_HbSliceState.eFault: // 故障相：码值锁存回放，仅复位沿出 [-] / fault, exit only on reset [-]
        ; // 锁存回放（R28） [-] / replay the latch only [-]
ELSE
    _iErr := 805; _eState := E_DL_HbSliceState.eFault; // 非法相位兜底 [-] / illegal phase fallback [-]
END_CASE

// 段 4｜限位钳位与出口映射（名实双出口，同源赋值）
IF rPos > fPosMaxMm THEN
    rPos := fPosMaxMm; // 上限位钳位 [mm] / clamp at the upper mechanical limit [mm]
END_IF
IF rPos < fPosMinMm THEN
    rPos := fPosMinMm; // 下限位钳位 [mm] / clamp at the lower mechanical limit [mm]
END_IF
eState := _eState; // 状态出口 [-] / state outlet [-]
rSlicePos := rPos; // 开度指令出口（已限位） [mm] / opening command outlet after limiting [mm]
iErrCode := _iErr; // 故障码出口（锁存值） [-] / error code outlet [-]
xReady := _eState = E_DL_HbSliceState.eReady; // 就绪位 = 就绪相镜像 [-] / ready mirrors the ready phase [-]
END_FUNCTION_BLOCK

(* ---- FB_DL_HeatExchangerFoulingTrend.st ---- *)
(*
  FB_DL_HeatExchangerFoulingTrend  —  换热器结垢趋势诊断（传热系数衰减速率） / Heat exchanger fouling trend diagnosis via UA decay rate
  分类 Category : DL_Process
  版本 Version  : 1.0.0
  来源 Source   : t1-2-oscat-building — 换热器族深化（与 HeatExchangerCtrl/HeatExchangerLmtd 分工：那两件管控制与 LMTD 计算，本件管结垢趋势诊断）
  溯源 Origin   : clean-room 实现，UA = 热负荷 / LMTD 为公开传热公式，未复制任何源码行
  功能 Function : 1) UA 估计：fUA := fHeatKw / fLmtdK（除法前域闸 fLmtdK >=
                  fLmtdMin 且 fHeatKw > 0，防除零与负商）；
                  2) 趋势窗：tTrendWin 单相独占 TON，窗内累计 UA 样本均值，
                  窗满判据 fUAavg < fUaRef × fUaTripPct / 100 → 039B 结垢
                  衰减超阈锁存（R190 归因唯一：判据无效走 039A，衰减超阈走 039B）；
                  3) 判据无效（LMTD 低于下限 / UA 非有限）→ ePause 相暂停采样
                  （双出口：判据恢复 / 撤使能，R98），判据无效为条件暂停不锁存；
                  4) 故障级：039A UA 换算非有限锁存（防御兜底）/ 039B 结垢衰减
                  超阈锁存 / 039C 组态非法 + ELSE 兜底归并；
                  5) 信息级三码：趋势窗采样完成 / 判据恢复 / 趋势复位（单拍沿）；
                  6) 解除式全当拍量（R240 落地），逐 BOOL 标注见段 4。
  边界 Boundary : ① 组态闸：fLmtdMin <= 0、fUaRef <= 0、fUaTripPct 不在
                  (0,100] 域、tTrendWin <= 0 → 039C 锁存，采样停发；
                  ② 非有限判据自反 + 差值自减双判（R79）；均值除法前判样本数
                  > 0（防除零）；
                  ③ 判据无效暂停为条件态不占故障码（R90 反证：暂停态由
                  bDtInvalid 镜像 + 相位出口可完整观测，不需加码）；
                  ④ 无 GVL 依赖：纯引脚输入输出，无外部变量引用，无物理 IO 地址。
  依赖 Depends  : Standard.library（TON / R_TRIG）
  码表 Error codes（Process 段 0005，窗口 039A~039C / 04C2~04C4）:
    16#0005_039A 故障级：UA 换算非有限锁存（防御兜底），锁存至 bReset
    16#0005_039B 故障级：结垢衰减超阈锁存（窗均 UA 低于 fUaTripPct 基准），锁存至 bReset
    16#0005_039C 故障级：组态非法（LMTD 下限/基准 UA/百分比/窗域非法）或相位落 ELSE 兜底（归并声明），锁存至 bReset
    16#0005_04C2 信息级：趋势窗采样完成沿（窗满判定拍）
    16#0005_04C3 信息级：判据恢复沿（ePause 恢复出口）
    16#0005_04C4 信息级：趋势复位沿（样本累计清零拍）
  修订历史 Revision :
    2026-11-19  v1.0.0  R42 首版（批次 3 · 序号 5）
*)

TYPE E_DL_HftState :
(
    eIdle   := 0,    // 未使能：不采样 / Idle, not sampling
    eRun    := 10,   // 采样中：UA 累计 / Run, UA accumulating
    ePause  := 20,   // 暂停：判据无效 / Pause, verdict invalid
    eFault  := 90    // 故障：非有限或超阈锁定 / Fault, latched
);
END_TYPE

FUNCTION_BLOCK FB_DL_HeatExchangerFoulingTrend
VAR_INPUT
    fHeatKw      : REAL := 0.0;       // 换热负荷 [kW]，调用方注入 / Heat duty
    fLmtdK       : REAL := 0.0;       // 对数平均温差 [K]，调用方注入（LMTD 属主为 HeatExchangerLmtd）/ LMTD
    fLmtdMin     : REAL := 1.0;       // LMTD 判据下限 [K]，域 > 0 / LMTD verdict minimum
    fUaRef       : REAL := 100.0;     // 洁净基准 UA [kW/K]，域 > 0 / Clean reference UA
    fUaTripPct   : REAL := 70.0;      // 结垢衰减跳闸百分比 [%]，域 (0,100] / Fouling trip percent
    tTrendWin    : TIME := T#60S;     // 趋势采样窗 [ms]，域 > 0 / Trend sampling window
    bTrendEn     : BOOL := FALSE;     // 趋势使能（电平）[-] / Trend enable, level
    bTrendRst    : BOOL := FALSE;     // 趋势复位指令，上升沿清样本累计 [-] / Trend reset command edge
    bReset       : BOOL := FALSE;     // 复位，上升沿清故障锁存 / Reset edge clears fault latch
END_VAR
VAR_OUTPUT
    eState       : E_DL_HftState;     // 状态出口，段尾单点映射 / State outlet
    fUaNow       : REAL;              // 当前 UA 估计 [kW/K] / Current UA estimate
    fUaWinAvg    : REAL;              // 趋势窗 UA 均值 [kW/K]（窗满刷新）/ Window UA average
    bVerdictBad  : BOOL;              // 判据无效镜像（ePause 相电平）[-] / Verdict-invalid mirror
    bError       : BOOL;              // 故障锁存标志 / Fault latch flag
    nErrId       : UDINT;             // 事件码，0 = 无事件 / Event code
END_VAR
VAR
    tonTrendWin  : TON;               // 趋势采样窗（单相独占），无条件刷新 / Trend window timer
    _eState      : E_DL_HftState := E_DL_HftState.eIdle;   // 内部相位，CASE 唯一写入目标 / Internal phase, the only CASE write target
    rtTrendRst   : R_TRIG;            // 趋势复位沿实例，无条件刷新 / Trend reset edge instance
    rtReset      : R_TRIG;            // 复位沿实例，无条件刷新 / Reset edge instance
    _fUa         : REAL;              // 逐拍 UA 估计 [kW/K]（当拍量）/ Per-scan UA estimate
    _bVerdictOk  : BOOL;              // 判据有效当拍量 [-] / Verdict-valid flag
    _bNonFin     : BOOL;              // UA 非有限当拍量 [-] / Non-finite UA flag
    _nSamples    : DINT;              // 窗内样本数 [个] / Sample count in window
    _fUaSum      : REAL;              // 窗内 UA 样本和 [kW/K] / UA sample sum in window
    _bFault      : BOOL;              // 故障锁存位（锁存量）/ Latched fault bit
    _uFault      : UDINT;             // 故障码锁存（锁存量）/ Latched fault code
    _uInfo       : UDINT;             // 信息码，每拍重算 / Transient info code
END_VAR

(* —— 段 0：定时器与沿实例无条件周期刷新（禁置于 IF/CASE 内） —— *)
_bVerdictOk := (fLmtdK >= fLmtdMin) AND (fHeatKw > 0.0);    // 判据有效（当拍量：分母域闸 + 正负荷）
IF _bVerdictOk THEN                  // 域内才做除法（防除零/防负商）
    _fUa := fHeatKw / fLmtdK;        // UA 估计（当拍量）
    _bNonFin := (_fUa <> _fUa) OR ((_fUa - _fUa) <> (_fUa - _fUa));
                                        // 非有限防御（NaN 自反 + 差值自减）
ELSE
    _fUa := 0.0;                     // 判据无效：UA 置 0（安全侧）
    _bNonFin := FALSE;               // 未做除法：非有限标志 FALSE
END_IF
rtTrendRst(CLK := bTrendRst);        // 趋势复位沿（每拍必调）
rtReset(CLK := bReset);              // 复位沿（每拍必调）
tonTrendWin(IN := (_eState = E_DL_HftState.eRun) AND _bVerdictOk, PT := tTrendWin);
                                        // 趋势窗（运行相 + 判据有效电平，暂停拍 IN 断）

(* —— 段 1：单拍量预清零（锁存量 _bFault/_uFault 与样本累计不入清单，禁同拍抹除） —— *)
_uInfo := 16#0000_0000;             // 信息码每拍重算
fUaNow := _fUa;                     // 当前 UA 出口（当拍量直出）
bVerdictBad := FALSE;               // 判据无效镜像缺省 FALSE
nErrId := 16#0000_0000;             // 事件码缺省无事件

(* —— 段 2：复位沿 + 组态域闸（判据当拍量） —— *)
IF rtReset.Q THEN                   // rtReset.Q = 当拍量
    _bFault := FALSE;               // 清故障锁存位
    _uFault := 16#0000_0000;        // 清故障锁存码
END_IF
IF (fLmtdMin <= 0.0) OR (fUaRef <= 0.0) OR (fUaTripPct <= 0.0) OR (fUaTripPct > 100.0)
   OR (TIME_TO_DINT(tTrendWin) <= 0) THEN
    _uFault := 16#0005_039C;        // 故障级：组态非法
    _bFault := TRUE;                // 故障标志与码位配对（R45）
END_IF
IF rtTrendRst.Q THEN                // 趋势复位沿（当拍量）
    _nSamples := 0;                 // 样本数清零
    _fUaSum := 0.0;                 // 样本和清零
    fUaWinAvg := 0.0;               // 窗均值清零
    _uInfo := 16#0005_04C4;         // 信息级：趋势复位沿
END_IF

(* —— 段 3：非有限锁存（判据当拍量） —— *)
IF _bNonFin THEN
    _uFault := 16#0005_039A;        // 故障级：UA 非有限（防御兜底）
    _bFault := TRUE;
END_IF

(* —— 段 4：故障解除式（R240 落地，逐 BOOL 标注）：
     rtReset.Q = 当拍量；NOT bTrendEn = 当拍量；_bVerdictOk = 当拍量。
     均不含锁存量（_bFault/_uFault），解除边真实可达（判据恢复 + 撤使能 + 复位沿）。 —— *)
IF rtReset.Q AND (NOT bTrendEn) AND _bVerdictOk AND (NOT _bNonFin) THEN
    _bFault := FALSE;               // 清故障锁存位（锁存量，仅此当拍量解除沿可清）
    _uFault := 16#0000_0000;        // 清故障锁存码（锁存量，仅本当拍量解除沿可清）
    IF _eState = E_DL_HftState.eFault THEN
        _eState := E_DL_HftState.eIdle;     // 故障相迁出：回未使能
    END_IF
END_IF

(* —— 段 5：相位机（CASE 全覆盖 + ELSE 兜底） —— *)
CASE _eState OF

E_DL_HftState.eIdle:
    IF bTrendEn AND (NOT _bFault) THEN
        _nSamples := 0;                 // 样本数清零（进相预置）
        _fUaSum := 0.0;                 // 样本和清零（进相预置）
        _eState := E_DL_HftState.eRun;  // 进采样相
    END_IF

E_DL_HftState.eRun:
    IF _bVerdictOk AND (NOT _bNonFin) THEN
        _fUaSum := _fUaSum + _fUa;      // 样本累计
        _nSamples := _nSamples + 1;     // 样本数递增
    ELSE
        _eState := E_DL_HftState.ePause;    // 判据无效：进暂停相
    END_IF
    IF tonTrendWin.Q THEN               // 窗满判定（单相独占 TON）
        IF _nSamples > 0 THEN           // 均值除法前判样本数（防除零）
            fUaWinAvg := _fUaSum / UDINT_TO_REAL(UDINT(_nSamples));    // 窗均值
        END_IF
        _uInfo := 16#0005_04C2;         // 信息级：趋势窗采样完成沿
        _nSamples := 0;                 // 窗重启：样本数清零
        _fUaSum := 0.0;                 // 窗重启：样本和清零
        IF fUaWinAvg < fUaRef * fUaTripPct / 100.0 THEN
            _uFault := 16#0005_039B;    // 故障级：结垢衰减超阈
            _bFault := TRUE;
        END_IF
    END_IF
    IF NOT bTrendEn THEN
        _eState := E_DL_HftState.eIdle; // 撤使能：回未使能相
    END_IF

E_DL_HftState.ePause:
    bVerdictBad := TRUE;                // 判据无效镜像（相电平）
    IF _bVerdictOk AND (NOT _bNonFin) THEN  // 出口 1：判据恢复（事件量）
        _uInfo := 16#0005_04C3;         // 信息级：判据恢复沿
        _eState := E_DL_HftState.eRun;  // 回采样相
    ELSIF NOT bTrendEn THEN             // 出口 2：撤使能（前置条件消失，R98 双出口）
        _eState := E_DL_HftState.eIdle; // 回未使能相
    END_IF

E_DL_HftState.eFault:
    ;                                   // 故障相：采样冻结，等解除沿（段 4 承载迁出）

ELSE
    _uFault := 16#0005_039C;            // 故障级：非法相位兜底（归并组态码，码表声明）
    _bFault := TRUE;
    _eState := E_DL_HftState.eFault;    // 强制回故障相

END_CASE

(* —— 段 6：出口单点映射（名实同源；锁存码回放，禁同拍抹除） —— *)
IF _bFault THEN
    nErrId := _uFault;              // 故障锁存码回放
    bVerdictBad := FALSE;           // 故障相判据镜像强制 FALSE
    fUaNow := 0.0;                  // 故障相 UA 出口强制 0（安全侧）
ELSE
    nErrId := _uInfo;               // 信息码
END_IF
bError := _bFault;                  // 故障标志与锁存位同源
eState := _eState;                  // 状态出口单点映射

END_FUNCTION_BLOCK

(* ---- FB_DL_HeatSealProfile.st ---- *)
(*
  FB_DL_HeatSealProfile  —  热封温度-压力-时间三参数配方曲线管理 / Heat-seal temperature-pressure-time profile
  分类 Category : DL_Process
  码位 Code     : 16#06_0_B0
  版本 Version  : 1.0.0
  来源 Source   : t2-7-packml — IEC 61131-3 标准语义的道莅防御性实现
  溯源 Origin   : clean-room 实现，PackML 热封段序公开语义借鉴，未复制任何源码行
                  （RESUME 承接 R36 §4 #15 规格；段推进语义对齐 FB_DL_StepSequencer，配方驻留对齐 FB_DL_RampSoakProfile，均不实例化）
  功能 Function : 1) 升温(Heat)→加压(Press)→冷却(Cool) 三段按配方时长推进（时长 0 的段跳过并记信息码）；
                  2) 各段实测温度/压力必须落在配方 ± 容差带内，越带记段不合格（_abSegBad 末段汇总 bProfileOk）；
                  3) 单段超 tSealMax 升级为 Fault；bAbort 在任意段立即进 Fault 并置 bReject。
  边界 Boundary : ① 配方时长为 0 的段跳过但记信息码；配方三段全为 0 判组态错不启动；
                  ② 容差/超时非法同判组态错；温度配方须为正值域（开尔文域防御）；
                  ③ bAbort 任意段立即进 Fault 并置 bReject（安全侧先撤输出）；
                  ④ CASE 全态覆盖 + ELSE 兜底（未知状态回 Idle 并置码，规格强制）；
                  ⑤ 解除式自证：bReject 解除 = bStart 上升沿 AND bReset（两引脚均可满足，R28-1）；
                  ⑥ 段判据 _abSegBad 为周期内锁存量，Done 相汇总后随新周期 bStart 上升沿清零。
  依赖 Depends  : 仅 Standard.library（TON/R_TRIG）；段序语义对齐 FB_DL_StepSequencer / FB_DL_RampSoakProfile（已注册，不实例化）
  码表 Error codes（本件格 06_0_B0，子码步进 +0x100）:
    16#0006_01B0 信息级：段时长为 0，该段跳过
    16#0006_02B0 故障级：组态非法（配方全 0 / 容差 <= 0 / tSealMax <= 0），锁存至复位
    16#0006_03B0 故障级：单段超时 tSealMax 升级
    16#0006_04B0 信息级：段参数越容差带（记段不合格）
    16#0006_05B0 信息级：中止判废（bAbort 触发）
    16#0006_06B0 故障级：状态机落 ELSE 兜底（非法相位 ID）

  修订历史 Revision :
    2026-11-18  v1.0.0  R38 首版
*)

TYPE E_DL_SealPhase :
(
    eIdle   := 0,    // 空闲：等启动指令 / Idle, waiting for start
    eHeat   := 10,   // 升温段 / Heating segment
    ePress  := 20,   // 加压段 / Pressing segment
    eCool   := 30,   // 冷却段 / Cooling segment
    eDone   := 40,   // 完成：曲线合格汇总落定 / Done, profile verdict settled
    eReject := 50,   // 判废：曲线不合格落定（非故障）/ Rejected, profile unfit
    eFault  := 90    // 故障：组态/超时/中止锁定 / Fault, latched
);
END_TYPE

FUNCTION_BLOCK FB_DL_HeatSealProfile
VAR_INPUT
    bStart         : BOOL := FALSE;              // 启动指令（上升沿）/ Start command
    bAbort         : BOOL := FALSE;              // 中止指令（任意段生效）/ Abort command
    bReset         : BOOL := FALSE;              // 复位（Fault/bReject 解除路径之一）/ Reset
    afSealTempC    : ARRAY[0..2] OF REAL;        // 配方温度三段 [°C] / Recipe temperatures
    afSealPressBar : ARRAY[0..2] OF REAL;        // 配方压力三段 [bar] / Recipe pressures
    atSealTimeMs   : ARRAY[0..2] OF TIME;        // 配方时长三段 [ms] / Recipe durations
    fTempActualC   : REAL := 0.0;                // 实测封口温度 [°C] / Actual seal temperature
    fPressActualBar: REAL := 0.0;                // 实测封口压力 [bar] / Actual seal pressure
    fTempTolC      : REAL := 5.0;                // 温度容差 [°C]，域 > 0 / Temperature tolerance
    fPressTolBar   : REAL := 0.5;                // 压力容差 [bar]，域 > 0 / Pressure tolerance
    tSealMax       : TIME := T#30S;              // 单段超时上限 [ms]，域 > 0 / Segment timeout ceiling
END_VAR
VAR_OUTPUT
    bSealing   : BOOL;                       // 封口进行中（Heat/Press/Cool 任一段）/ Sealing in progress
    bProfileOk : BOOL;                       // 曲线合格（末段汇总）/ Profile verdict
    bReject    : BOOL;                       // 判废锁存（解除式：bStart 沿 AND bReset）/ Reject latch
    nSegment   : INT;                        // 当前段号 [0..2] / Current segment index
    fElapsedMs : REAL;                       // 当前段已走时长 [ms] / Segment elapsed time
    nErrId     : UDINT;                      // 事件码，0 = 无事件 / Event code
    eState     : E_DL_SealPhase;             // 状态出口，段尾单点映射 / State outlet
END_VAR
VAR
    tonSeg     : TON;                        // 当前段配方时长计时，段 0 无条件刷新 / Segment recipe timer
    tonSegMax  : TON;                        // 单段超时计时，段 0 无条件刷新 / Segment timeout timer
    tonFaultWch: TON;                        // 故障观察窗，自复位 / Fault watch window, self-resetting
    rtStart    : R_TRIG;                     // 启动上升沿 / Start rising edge
    rtReset    : R_TRIG;                     // 复位上升沿 / Reset rising edge
    _eState    : E_DL_SealPhase := E_DL_SealPhase.eIdle;   // 内部相位（CASE 唯一写入目标）/ Internal phase
    _nSeg      : INT;                        // 当前段号内部量 [0..2] / Internal segment index
    _abSegBad  : ARRAY[0..2] OF BOOL;        // 段不合格锁存（越带记段）/ Per-segment unfit latch
    _bAnyBad   : BOOL;                       // 任一段不合格聚合 / Any segment unfit aggregate
    _bSkip     : BOOL;                       // 段时长为 0 跳过标志（本拍重算）/ Zero-duration skip flag
    _uFault    : UDINT;                      // 故障码锁存 / Latched fault code
    _uInfo     : UDINT;                      // 信息码，每拍重算 / Info code
    _bFault    : BOOL;                       // 故障锁存位 / Latched fault bit
    _bCfgBad   : BOOL;                       // 组态非法聚合 / Configuration invalid aggregate
    _bRejectL  : BOOL;                       // 判废锁存保持量 / Reject latch held quantity
    _nK        : INT;                        // 循环计数器 / Loop counter
END_VAR
VAR CONSTANT
    DL_WatchPt : TIME := T#2S;   // 故障观察窗 [ms]，自复位 / Fault watch window
END_VAR

(* —— 段 0：定时器与边沿无条件周期刷新（R182：调用语句不得置于 IF/CASE 内） —— *)
rtStart(CLK := bStart);                                          // 启动上升沿，每拍必调
rtReset(CLK := bReset);                                          // 复位上升沿，每拍必调
tonFaultWch(IN := (NOT tonFaultWch.Q), PT := DL_WatchPt);        // 观察窗自复位（表达式入参）
tonSeg(IN := (_eState = E_DL_SealPhase.eHeat) OR (_eState = E_DL_SealPhase.ePress)
            OR (_eState = E_DL_SealPhase.eCool), PT := atSealTimeMs[_nSeg]);   // 段配方时长（表达式入参）
tonSegMax(IN := (_eState = E_DL_SealPhase.eHeat) OR (_eState = E_DL_SealPhase.ePress)
              OR (_eState = E_DL_SealPhase.eCool), PT := tSealMax);   // 单段超时（表达式入参）

(* —— 段 1：单拍量预清零（锁存量 _uFault/_bFault/_bRejectL/_abSegBad/_bAnyBad 不入清单，R187①） —— *)
_uInfo := 16#0000_0000;         // 信息码每拍重算
bSealing := FALSE;              // 封口出口缺省 FALSE（段 8 单点置位）
_bCfgBad := FALSE;              // 组态非法预清零
_bSkip := FALSE;                // 跳过标志预清零
nErrId := 16#0000_0000;         // 事件码缺省无事件

(* —— 段 2：组态域闸（覆盖全部参与判据换算的引脚，R151） —— *)
IF (fTempTolC <= 0.0) OR (fPressTolBar <= 0.0) OR (TIME_TO_DINT(tSealMax) <= 0) THEN
    _bCfgBad := TRUE;           // 容差/超时非法
END_IF
FOR _nK := 0 TO 2 DO
    IF (afSealTempC[_nK] <> afSealTempC[_nK]) OR (afSealTempC[_nK] <= 0.0)
       OR (afSealTempC[_nK] > 400.0) THEN
        _bCfgBad := TRUE;       // 温度配方非法（正值域，开尔文域防御）
    END_IF
    IF (afSealPressBar[_nK] <> afSealPressBar[_nK]) OR (afSealPressBar[_nK] <= 0.0)
       OR (afSealPressBar[_nK] > 10.0) THEN
        _bCfgBad := TRUE;       // 压力配方非法（正值域上限防御）
    END_IF
END_FOR
IF (TIME_TO_DINT(atSealTimeMs[0]) <= 0) AND (TIME_TO_DINT(atSealTimeMs[1]) <= 0)
   AND (TIME_TO_DINT(atSealTimeMs[2]) <= 0) THEN
    _bCfgBad := TRUE;           // 配方三段全 0：不启动（规格强制）
END_IF

(* —— 段 3：复位沿（bReject 解除式：bStart 上升沿 AND bReset；Fault 解除 = bReset） —— *)
IF rtReset.Q THEN
    IF rtStart.Q THEN
        _bRejectL := FALSE;     // 判废锁存清零（解除式自证路径）
    END_IF
    _bFault := FALSE;           // 清故障锁存位
    _uFault := 16#0000_0000;
    IF _eState = E_DL_SealPhase.eFault THEN
        _eState := E_DL_SealPhase.eIdle;    // 故障相回空闲
    END_IF
END_IF

(* —— 段 4：中止拦截（任意段立即升级，安全侧先撤输出——出口由 Fault 相缺省保证） —— *)
IF bAbort AND (_eState <> E_DL_SealPhase.eIdle) AND (_eState <> E_DL_SealPhase.eFault)
   AND (_eState <> E_DL_SealPhase.eDone) AND (_eState <> E_DL_SealPhase.eReject) THEN
    _uFault := 16#0006_03B0;    // 中止按故障级升级（撤输出）
    _bFault := TRUE;            // 锁存
    _bRejectL := TRUE;          // 判废锁存（bAbort 置 bReject，规格强制）
    _uInfo := 16#0006_05B0;     // 信息级：中止判废
    _eState := E_DL_SealPhase.eFault;
END_IF

(* —— 段 5：相位机（只做迁移与判据记账；出口在段 8） —— *)
CASE _eState OF

E_DL_SealPhase.eIdle:
    IF _bCfgBad THEN
        _uFault := 16#0006_02B0;            // 故障级：组态非法
        _bFault := TRUE;                    // 锁存（复位沿可清）
        _eState := E_DL_SealPhase.eFault;
    ELSIF rtStart.Q THEN
        _nSeg := 0;                         // 段号归零
        FOR _nK := 0 TO 2 DO
            _abSegBad[_nK] := FALSE;        // 段判据清零（新周期）
        END_FOR
        _bAnyBad := FALSE;                  // 聚合清零
        bProfileOk := FALSE;                // 曲线结论复位（Done 相重判）
        _eState := E_DL_SealPhase.eHeat;    // 进升温段
    END_IF

E_DL_SealPhase.eHeat:
    IF TIME_TO_DINT(atSealTimeMs[_nSeg]) <= 0 THEN
        _bSkip := TRUE;                     // 段时长为 0：跳过
        _uInfo := 16#0006_01B0;             // 信息级：段跳过
        _nSeg := _nSeg + 1;                 // 段号递增（上限守卫在 CASE 前判）
        IF _nSeg > 2 THEN
            _eState := E_DL_SealPhase.eDone;    // 三段走完：进完成相
        ELSE
            _eState := E_DL_SealPhase.ePress;   // 进加压段
        END_IF
    ELSIF tonSeg.Q THEN
        IF ABS(fTempActualC - afSealTempC[_nSeg]) > fTempTolC THEN
            _abSegBad[_nSeg] := TRUE;       // 越温带：记段不合格
            _uInfo := 16#0006_04B0;         // 信息级：段越带
        END_IF
        _nSeg := _nSeg + 1;
        IF _nSeg > 2 THEN
            _eState := E_DL_SealPhase.eDone;
        ELSE
            _eState := E_DL_SealPhase.ePress;
        END_IF
    ELSIF tonSegMax.Q THEN
        _uFault := 16#0006_03B0;            // 故障级：单段超时升级
        _bFault := TRUE;
        _eState := E_DL_SealPhase.eFault;
    END_IF

E_DL_SealPhase.ePress:
    IF TIME_TO_DINT(atSealTimeMs[_nSeg]) <= 0 THEN
        _bSkip := TRUE;
        _uInfo := 16#0006_01B0;
        _nSeg := _nSeg + 1;
        IF _nSeg > 2 THEN
            _eState := E_DL_SealPhase.eDone;
        ELSE
            _eState := E_DL_SealPhase.eCool;
        END_IF
    ELSIF tonSeg.Q THEN
        IF ABS(fTempActualC - afSealTempC[_nSeg]) > fTempTolC THEN
            _abSegBad[_nSeg] := TRUE;
            _uInfo := 16#0006_04B0;
        END_IF
        IF ABS(fPressActualBar - afSealPressBar[_nSeg]) > fPressTolBar THEN
            _abSegBad[_nSeg] := TRUE;       // 越压带：记段不合格
            _uInfo := 16#0006_04B0;
        END_IF
        _nSeg := _nSeg + 1;
        IF _nSeg > 2 THEN
            _eState := E_DL_SealPhase.eDone;
        ELSE
            _eState := E_DL_SealPhase.eCool;
        END_IF
    ELSIF tonSegMax.Q THEN
        _uFault := 16#0006_03B0;
        _bFault := TRUE;
        _eState := E_DL_SealPhase.eFault;
    END_IF

E_DL_SealPhase.eCool:
    IF TIME_TO_DINT(atSealTimeMs[_nSeg]) <= 0 THEN
        _bSkip := TRUE;
        _uInfo := 16#0006_01B0;
        _nSeg := _nSeg + 1;
        _eState := E_DL_SealPhase.eDone;    // 冷却为末段：进完成相
    ELSIF tonSeg.Q THEN
        IF ABS(fTempActualC - afSealTempC[_nSeg]) > fTempTolC THEN
            _abSegBad[_nSeg] := TRUE;
            _uInfo := 16#0006_04B0;
        END_IF
        _nSeg := _nSeg + 1;
        _eState := E_DL_SealPhase.eDone;
    ELSIF tonSegMax.Q THEN
        _uFault := 16#0006_03B0;
        _bFault := TRUE;
        _eState := E_DL_SealPhase.eFault;
    END_IF

E_DL_SealPhase.eDone:
    _bAnyBad := _abSegBad[0] OR _abSegBad[1] OR _abSegBad[2];   // 末段汇总
    bProfileOk := NOT _bAnyBad;             // 曲线合格结论
    IF _bAnyBad THEN
        _bRejectL := TRUE;                  // 不合格判废
    END_IF
    IF NOT bStart THEN
        _eState := E_DL_SealPhase.eIdle;    // 指令撤销：回空闲（结论保持）
    END_IF

E_DL_SealPhase.eReject:
    ;                                       // 预留相（判废经 Done 落定，本相不进入——保留枚举全态覆盖）

E_DL_SealPhase.eFault:
    ;                                       // 故障相：等复位沿（段 3 承载解除）

ELSE
    _uFault := 16#0006_06B0;                // 故障级：非法相位 ID 兜底
    _bFault := TRUE;                        // 锁存
    _eState := E_DL_SealPhase.eIdle;        // 未知状态回 Idle（规格强制）

END_CASE

(* —— 段 6：出口单点映射（名实同源；锁存码回放，禁同拍抹除） —— *)
bSealing := (_eState = E_DL_SealPhase.eHeat) OR (_eState = E_DL_SealPhase.ePress)
            OR (_eState = E_DL_SealPhase.eCool);            // 封口出口：三段任一
nSegment := _nSeg;                          // 段号出口
fElapsedMs := TIME_TO_REAL(tonSegMax.ET);   // 已走时长出口（超时窗实时值 [ms]）
bReject := _bRejectL;                       // 判废出口 = 锁存量（置位同拍不被抹）
IF _bFault THEN
    nErrId := _uFault;          // 故障锁存码回放
    bSealing := FALSE;          // 故障相封口出口强制 FALSE（安全侧）
ELSE
    nErrId := _uInfo;           // 信息码
END_IF
eState := _eState;              // 状态出口单点映射

END_FUNCTION_BLOCK
